(* IEC 61131-3 sources: TetherPLC/compat/tc3 (part 2) *)

(* ---- tc3_analytics.st ---- *)
// tc3_analytics.st — Tc3_Analytics surface (TF3510/TF3500/TF3520):
// measurement analytics.  TwinCAT's full library is ~670 APIs
// behind a licensed analytics engine; the local measurement-side
// primitives (event counting, windowed statistics, sample
// logging) are pure-ST here and fully functional, while the
// engine-backed surfaces (storage provider, MQTT/HTTP egress
// transport) report an honest engine-absent error.
//
// Differences from the TwinCAT library
// (docs/plc/compat/README.md):
//   - TwinCAT's class/method/object model is flattened into
//     FB_* blocks with Execute-style inputs, matching the other
//     TetherPLC compat surfaces.
//   - The ring logger exposes the newest N samples via indexed
//     outputs Slot0..Slot7 plus Count; a real circular-buffer
//     API needs dynamic memory we do not model.
//   - Storage/provider and transport FBs accept the command,
//     run a bounded handshake, then fail ErrorId=1
//     (engine-unavailable): no database or MQTT egress is faked.

// ---- FB_AnalyticsCounter: edge counter + rate per window ----
FUNCTION_BLOCK FB_AnalyticsCounter
VAR_INPUT
    Enable : BOOL;
    Event : BOOL;               // count rising edges
    WindowTime : LREAL;         // seconds per rate window
    CycleTime : LREAL;          // task cycle seconds
    Reset : BOOL;
END_VAR
VAR_OUTPUT
    Total : UDINT;
    WindowCount : UDINT;
    Rate : LREAL;               // events per second (last window)
    WindowDone : BOOL;
END_VAR
VAR
    prev : BOOL;
    acc : LREAL;
END_VAR
    WindowDone := FALSE;
    IF Reset THEN
        Total := 0;
        WindowCount := 0;
        Rate := 0.0;
        acc := 0.0;
        prev := FALSE;
    END_IF;
    IF NOT Enable THEN
        prev := Event;
        RETURN;
    END_IF;
    IF Event AND NOT prev THEN
        Total := Total + 1;
        WindowCount := WindowCount + 1;
    END_IF;
    prev := Event;
    acc := acc + CycleTime;
    IF WindowTime > 0.0 AND acc >= WindowTime THEN
        Rate := UDINT_TO_LREAL(WindowCount) / acc;
        WindowCount := 0;
        acc := 0.0;
        WindowDone := TRUE;
    END_IF;
END_FUNCTION_BLOCK

// ---- FB_AnalyticsStats: running + windowed min/max/mean ----
FUNCTION_BLOCK FB_AnalyticsStats
VAR_INPUT
    Execute : BOOL;             // sample the input when TRUE
    Sample : LREAL;
    Clear : BOOL;
END_VAR
VAR_OUTPUT
    Count : UDINT;
    Min : LREAL;
    Max : LREAL;
    Mean : LREAL;
    Valid : BOOL;
END_VAR
VAR
    sum : LREAL;
END_VAR
    Valid := FALSE;
    IF Clear THEN
        Count := 0;
        Min := 0.0;
        Max := 0.0;
        Mean := 0.0;
        sum := 0.0;
    END_IF;
    IF NOT Execute THEN RETURN; END_IF;
    IF Count = 0 THEN
        Min := Sample;
        Max := Sample;
    ELSE
        IF Sample < Min THEN Min := Sample; END_IF;
        IF Sample > Max THEN Max := Sample; END_IF;
    END_IF;
    Count := Count + 1;
    sum := sum + Sample;
    Mean := sum / UDINT_TO_LREAL(Count);
    Valid := TRUE;
END_FUNCTION_BLOCK

// ---- FB_AnalyticsLogger: 8-deep ring of timestamped samples ----
FUNCTION_BLOCK FB_AnalyticsLogger
VAR_INPUT
    Record : BOOL;              // rising edge stores a sample
    Value : LREAL;
    Timestamp : LREAL;          // caller-supplied time tag
    Clear : BOOL;
END_VAR
VAR_OUTPUT
    Count : UDINT;              // total records stored
    Slot0 : LREAL; Slot1 : LREAL; Slot2 : LREAL; Slot3 : LREAL;
    Slot4 : LREAL; Slot5 : LREAL; Slot6 : LREAL; Slot7 : LREAL;
    LastTs : LREAL;
    Overflow : BOOL;            // wrapped at least once
END_VAR
VAR
    head : UDINT;
    prev : BOOL;
END_VAR
    IF Clear THEN
        Count := 0;
        head := 0;
        LastTs := 0.0;
        Overflow := FALSE;
        Slot0 := 0.0; Slot1 := 0.0; Slot2 := 0.0; Slot3 := 0.0;
        Slot4 := 0.0; Slot5 := 0.0; Slot6 := 0.0; Slot7 := 0.0;
    END_IF;
    IF Record AND NOT prev THEN
        IF head = 0 THEN Slot0 := Value; END_IF;
        IF head = 1 THEN Slot1 := Value; END_IF;
        IF head = 2 THEN Slot2 := Value; END_IF;
        IF head = 3 THEN Slot3 := Value; END_IF;
        IF head = 4 THEN Slot4 := Value; END_IF;
        IF head = 5 THEN Slot5 := Value; END_IF;
        IF head = 6 THEN Slot6 := Value; END_IF;
        IF head = 7 THEN Slot7 := Value; END_IF;
        head := head + 1;
        IF head >= 8 THEN
            head := 0;
            Overflow := TRUE;
        END_IF;
        Count := Count + 1;
        LastTs := Timestamp;
    END_IF;
    prev := Record;
END_FUNCTION_BLOCK

// ---- FB_AnalyticsStore: engine-backed storage provider ----
// Honest engine-absent block: accepts a flush/store command,
// holds Busy for a bounded handshake, then fails with
// ErrorId=1 — no database write is ever claimed.
FUNCTION_BLOCK FB_AnalyticsStore
VAR_INPUT
    Execute : BOOL;
    Abort : BOOL;
    ProviderPath : STRING;      // e.g. database/Influx endpoint
    RecordCount : UDINT;
END_VAR
VAR_OUTPUT
    Busy : BOOL;
    Error : BOOL;
    ErrorId : UDINT;            // 0 none, 1 engine-unavailable,
                                // 2 bad-provider, 3 aborted
    Done : BOOL;
END_VAR
VAR
    phase : INT;
    tmo : UDINT;
END_VAR
    Done := FALSE;
    IF phase = 0 THEN
        Busy := FALSE;
        IF Execute THEN
            Busy := TRUE;
            Error := FALSE;
            ErrorId := 0;
            tmo := 0;
            IF ProviderPath = '' THEN
                Error := TRUE;
                ErrorId := 2;
                phase := 2;
            ELSE
                phase := 1;
            END_IF;
        END_IF;
    ELSIF phase = 1 THEN
        tmo := tmo + 1;
        IF tmo >= 4 THEN
            Busy := FALSE;
            Error := TRUE;
            ErrorId := 1;       // engine-unavailable
            phase := 2;
        END_IF;
    ELSE
        Busy := FALSE;
        IF NOT Execute THEN phase := 0; END_IF;
    END_IF;
    IF Abort AND phase = 1 THEN
        Busy := FALSE;
        Error := TRUE;
        ErrorId := 3;
        phase := 2;
    END_IF;
    Done := (phase = 2);
END_FUNCTION_BLOCK

(* ---- tc3_ba_common.st ---- *)
// tc3_ba_common.st — Tc3_BA_Common + Tc3_BA2_Common surface
// (TwinCAT_3_PLC_Lib_Tc3_BA*_Common_EN): pure-ST building-
// automation commons — time-of-day helpers, edge/COV triggers,
// ramp limiters, 2-point switches, PID, sequence controller,
// and a bounded dynamic array.  KL32xx terminal config is not
// modeled (blocks take scaled process values).
//
// Differences: the BA_* enum-validity helpers map to plain
// range checks (enums are INT here); the DynamicArray is a
// bounded fixed-capacity variant (no heap growth).

// ---- F_BA_RemMsTp: ms remaining to a target time ----
FUNCTION F_BA_RemMsTp : UDINT
VAR_INPUT
    tNow : UDINT;               // ms
    tTarget : UDINT;
END_VAR
    IF tTarget >= tNow THEN
        F_BA_RemMsTp := tTarget - tNow;
    ELSE
        F_BA_RemMsTp := 0;
    END_IF;
END_FUNCTION

// ---- F_BA_RemSecsTp: s remaining to a target ----
FUNCTION F_BA_RemSecsTp : UDINT
VAR_INPUT
    tNow : UDINT;
    tTarget : UDINT;
END_VAR
    IF tTarget >= tNow THEN
        F_BA_RemSecsTp := tTarget - tNow;
    ELSE
        F_BA_RemSecsTp := 0;
    END_IF;
END_FUNCTION

// ---- F_BA_IsWeekdayValid: 1..7 range check ----
FUNCTION F_BA_IsWeekdayValid : BOOL
VAR_INPUT
    day : INT;
END_VAR
    F_BA_IsWeekdayValid := day >= 1 AND day <= 7;
END_FUNCTION

// ---- F_BA_IsUnitValid: unit-id range check ----
FUNCTION F_BA_IsUnitValid : BOOL
VAR_INPUT
    unit : INT;
END_VAR
    F_BA_IsUnitValid := unit >= 0 AND unit <= 255;
END_FUNCTION

// ---- FB_BA_RFTrig: rising/falling edge detector ----
FUNCTION_BLOCK FB_BA_RFTrig
VAR_INPUT
    bIn : BOOL;
END_VAR
VAR_OUTPUT
    bRise : BOOL;
    bFall : BOOL;
END_VAR
VAR
    prev : BOOL;
END_VAR
    bRise := bIn AND NOT prev;
    bFall := NOT bIn AND prev;
    prev := bIn;
END_FUNCTION_BLOCK

// ---- FB_BA_ATrigCOV: change-of-value trigger ----
// Fires when the input changes by more than fDelta since the
// last reported value.
FUNCTION_BLOCK FB_BA_ATrigCOV
VAR_INPUT
    bEnable : BOOL;
    fIn : LREAL;
    fDelta : LREAL;
END_VAR
VAR_OUTPUT
    bTrig : BOOL;
    fOut : LREAL;
END_VAR
VAR
    fLast : LREAL;
    init : BOOL;
END_VAR
    bTrig := FALSE;
    IF NOT bEnable THEN init := FALSE; RETURN; END_IF;
    IF NOT init THEN
        fLast := fIn;
        init := TRUE;
        bTrig := TRUE;
        fOut := fIn;
        RETURN;
    END_IF;
    IF fIn - fLast >= fDelta OR fLast - fIn >= fDelta THEN
        fLast := fIn;
        fOut := fIn;
        bTrig := TRUE;
    END_IF;
END_FUNCTION_BLOCK

// ---- FB_BA_RampLmt: ramp with output clamp ----
FUNCTION_BLOCK FB_BA_RampLmt
VAR_INPUT
    bEnable : BOOL;
    fIn : LREAL;
    fSlewUp : LREAL;            // unit/s
    fSlewDown : LREAL;
    fMin : LREAL;
    fMax : LREAL;
    CycleTime : LREAL;
END_VAR
VAR_OUTPUT
    fOut : LREAL;
    bAtTarget : BOOL;
END_VAR
    IF NOT bEnable THEN bAtTarget := FALSE; RETURN; END_IF;
    IF fOut < fIn THEN
        fOut := fOut + fSlewUp * CycleTime;
        IF fOut > fIn THEN fOut := fIn; END_IF;
    ELSIF fOut > fIn THEN
        fOut := fOut - fSlewDown * CycleTime;
        IF fOut < fIn THEN fOut := fIn; END_IF;
    END_IF;
    IF fOut > fMax THEN fOut := fMax; END_IF;
    IF fOut < fMin THEN fOut := fMin; END_IF;
    bAtTarget := fOut = fIn;
END_FUNCTION_BLOCK

// ---- FB_BA_Swi2P: two-point switch ----
FUNCTION_BLOCK FB_BA_Swi2P
VAR_INPUT
    bEnable : BOOL;
    fIn : LREAL;
    fOn : LREAL;
    fOff : LREAL;
END_VAR
VAR_OUTPUT
    bOut : BOOL;
END_VAR
VAR
    q : BOOL;
END_VAR
    IF NOT bEnable THEN q := FALSE; bOut := FALSE; RETURN; END_IF;
    IF fIn >= fOn THEN q := TRUE; END_IF;
    IF fIn <= fOff THEN q := FALSE; END_IF;
    bOut := q;
END_FUNCTION_BLOCK

// ---- FB_BA_SwiHys2P: two-point switch with hysteresis ----
FUNCTION_BLOCK FB_BA_SwiHys2P
VAR_INPUT
    bEnable : BOOL;
    fIn : LREAL;
    fSp : LREAL;
    fHys : LREAL;
    bInvert : BOOL;
END_VAR
VAR_OUTPUT
    bOut : BOOL;
END_VAR
VAR
    q : BOOL;
END_VAR
    IF NOT bEnable THEN q := FALSE; bOut := FALSE; RETURN; END_IF;
    IF bInvert THEN
        IF fIn >= fSp + fHys THEN q := TRUE; END_IF;
        IF fIn <= fSp THEN q := FALSE; END_IF;
    ELSE
        IF fIn <= fSp - fHys THEN q := TRUE; END_IF;
        IF fIn >= fSp THEN q := FALSE; END_IF;
    END_IF;
    bOut := q;
END_FUNCTION_BLOCK

// ---- FB_BA_PIDCtrl: PI controller with anti-windup ----
FUNCTION_BLOCK FB_BA_PIDCtrl
VAR_INPUT
    bEnable : BOOL;
    fActual : LREAL;
    fSetpoint : LREAL;
    fKp : LREAL;
    fTi : LREAL;                // s; 0 = P only
    fOutMin : LREAL;
    fOutMax : LREAL;
    CycleTime : LREAL;
END_VAR
VAR_OUTPUT
    fOut : LREAL;
    fError : LREAL;
END_VAR
VAR
    iTerm : LREAL;
END_VAR
    IF NOT bEnable THEN
        fOut := fOutMin; iTerm := 0.0; fError := 0.0;
        RETURN;
    END_IF;
    fError := fSetpoint - fActual;
    iTerm := iTerm + fError * CycleTime;
    fOut := fKp * fError;
    IF fTi > 0.0 THEN
        fOut := fKp * (fError + iTerm / fTi);
    END_IF;
    IF fOut > fOutMax THEN
        fOut := fOutMax;
        iTerm := iTerm - fError * CycleTime;
    END_IF;
    IF fOut < fOutMin THEN
        fOut := fOutMin;
        iTerm := iTerm - fError * CycleTime;
    END_IF;
END_FUNCTION_BLOCK

// ---- FB_BA_SeqCtrl: sequence controller ----
// Distributes a 0..100 demand across up to 4 sequential
// stages (each stage gets a slice of the demand range).
FUNCTION_BLOCK FB_BA_SeqCtrl
VAR_INPUT
    bEnable : BOOL;
    fDemand : LREAL;            // 0..100 %
    nStages : INT;              // 1..4
END_VAR
VAR_OUTPUT
    fStage1 : LREAL;            // each 0..100
    fStage2 : LREAL;
    fStage3 : LREAL;
    fStage4 : LREAL;
END_VAR
VAR
    seg : LREAL;
    rem : LREAL;
    nR : LREAL;
END_VAR
    IF NOT bEnable OR nStages <= 0 THEN
        fStage1 := 0.0; fStage2 := 0.0;
        fStage3 := 0.0; fStage4 := 0.0;
        RETURN;
    END_IF;
    nR := DINT_TO_LREAL(INT_TO_DINT(nStages));
    seg := 100.0 / nR;
    rem := fDemand;
    fStage1 := rem; IF fStage1 > seg THEN fStage1 := seg; END_IF;
    IF fStage1 < 0.0 THEN fStage1 := 0.0; END_IF;
    rem := rem - seg;
    fStage2 := rem; IF fStage2 > seg THEN fStage2 := seg; END_IF;
    IF fStage2 < 0.0 THEN fStage2 := 0.0; END_IF;
    rem := rem - seg;
    fStage3 := rem; IF fStage3 > seg THEN fStage3 := seg; END_IF;
    IF fStage3 < 0.0 THEN fStage3 := 0.0; END_IF;
    rem := rem - seg;
    fStage4 := rem; IF fStage4 > seg THEN fStage4 := seg; END_IF;
    IF fStage4 < 0.0 THEN fStage4 := 0.0; END_IF;
    // normalize each stage to 0..100 of its own slice
    fStage1 := fStage1 * 100.0 / seg;
    fStage2 := fStage2 * 100.0 / seg;
    fStage3 := fStage3 * 100.0 / seg;
    fStage4 := fStage4 * 100.0 / seg;
END_FUNCTION_BLOCK

// ---- FB_BA_DynamicArray: bounded key->value store ----
// Fixed capacity 16; key 0 is empty.
FUNCTION_BLOCK FB_BA_DynamicArray
VAR_INPUT
    bEnable : BOOL;
    Op : INT;                   // 1=set, 2=get, 3=remove, 4=find
    Key : UDINT;
    Value : LREAL;
END_VAR
VAR_OUTPUT
    Done : BOOL;
    Found : BOOL;
    OutValue : LREAL;
    Count : INT;
    Free : INT;
END_VAR
VAR
    keys : ARRAY[0..15] OF UDINT;
    vals : ARRAY[0..15] OF LREAL;
    cnt : INT;
    i : INT;
    slot : INT;
END_VAR
    Done := FALSE;
    Found := FALSE;
    OutValue := 0.0;
    IF NOT bEnable THEN RETURN; END_IF;
    slot := -1;
    FOR i := 0 TO 15 DO
        IF keys[i] = Key THEN slot := i; END_IF;
    END_FOR;
    IF Op = 1 THEN
        IF slot >= 0 THEN
            vals[slot] := Value;
            Found := TRUE;
            Done := TRUE;
        ELSE
            FOR i := 0 TO 15 DO
                IF slot < 0 AND keys[i] = 0 THEN slot := i; END_IF;
            END_FOR;
            IF slot >= 0 THEN
                keys[slot] := Key;
                vals[slot] := Value;
                cnt := cnt + 1;
                Done := TRUE;
            END_IF;
        END_IF;
    ELSIF Op = 2 OR Op = 4 THEN
        IF slot >= 0 THEN
            Found := TRUE;
            Done := TRUE;
            OutValue := vals[slot];
        END_IF;
    ELSIF Op = 3 THEN
        IF slot >= 0 THEN
            keys[slot] := 0;
            vals[slot] := 0.0;
            cnt := cnt - 1;
            Found := TRUE;
            Done := TRUE;
        END_IF;
    END_IF;
    Count := cnt;
    Free := 16 - cnt;
END_FUNCTION_BLOCK

(* ---- tc3_bacnet.st ---- *)
// Tc3_sACN -> Tc3_BACnetRev14 BACnet/IP client wrappers.
// Beckhoff's BACnet integration is device-configuration-driven
// (FBs are generated per configured device in TwinCAT), so there
// is no static TwinCAT FB API to mirror; these wrappers expose
// the tplc-bacnet service (ASHRAE 135 over UDP 47808) as
// poll-driven function blocks in the same shape as the other
// compat libraries.
// Differences from a TwinCAT BACnet device binding, documented in
// docs/plc/compat/README.md:
//   - Who-Is/ReadProperty/WriteProperty only; no COV subscriptions,
//     no device-object discovery beyond I-Am fields, no segmentation.
//   - Values cross as raw BACnet application-tag payload bytes:
//     nValueType selects the tag (1=boolean, 2=unsigned, 3=integer,
//     4=real, 5=double, 6=octetString, 7=characterString,
//     9=enumerated, 12=objectIdentifier) and pValue holds the tag
//     payload in wire byte order.
//   - nErrId carries tplc-bacnet service/transport codes.
// Sources: docs/plc/plan/21-twincat-libraries.md §7 (TF8020).

FUNCTION_BLOCK FB_BACnet_WhoIs
VAR_INPUT
    sHost : STRING[15];        // "" or "255.255.255.255" = broadcast
    nPort : UDINT := 47808;
    bHasRange : BOOL;
    nRangeLo : UDINT;
    nRangeHi : UDINT;
    bExecute : BOOL;
    tTimeout : TIME := T#1S;
END_VAR
VAR_OUTPUT
    bBusy : BOOL;
    bDone : BOOL;
    bError : BOOL;
    nErrId : UDINT;
    nStatus : DINT;
    nDevCount : UDINT;
    nDevId : ARRAY[0..7] OF UDINT;   // (objType<<22)|instance
    nDevIp : ARRAY[0..31] OF BYTE;   // 4 bytes per device
    nDevVendor : UDINT;
    nDevMaxApdu : UDINT;
    nDevSeg : UDINT;
END_VAR
VAR
    bac : FB_Bacnet;
    i : UDINT;
END_VAR
    bac.FUNC := 1;
    bac.HOST := sHost;
    bac.PORT := nPort;
    bac.HAS_RANGE := bHasRange;
    bac.RANGE_LO := nRangeLo;
    bac.RANGE_HI := nRangeHi;
    bac.TIMEOUT := tTimeout;
    bac.EXEC := bExecute;
    bac();
    bBusy := bac.BUSY;
    bDone := bac.DONE;
    nStatus := bac.STATUS;
    nErrId := bac.ERRID;
    nDevCount := bac.DEV_COUNT;
    nDevVendor := bac.DEV_VENDOR;
    nDevMaxApdu := bac.DEV_MAX_APDU;
    nDevSeg := bac.DEV_SEG;
    IF bac.DONE THEN
        i := 0;
        WHILE i < bac.DEV_COUNT AND i < 8 DO
            nDevId[i] := bac.DEV_ID[i];
            nDevIp[i*4] := bac.DEV_IP[i*4];
            nDevIp[i*4+1] := bac.DEV_IP[i*4+1];
            nDevIp[i*4+2] := bac.DEV_IP[i*4+2];
            nDevIp[i*4+3] := bac.DEV_IP[i*4+3];
            i := i + 1;
        END_WHILE;
    END_IF;
    bError := (bac.ERRID <> 0) OR (bac.STATUS >= 2);
END_FUNCTION_BLOCK

FUNCTION_BLOCK FB_BACnet_ReadProperty
VAR_INPUT
    sHost : STRING[15];
    nPort : UDINT := 47808;
    nObjType : UDINT;          // e.g. 8=device, 0=analogInput
    nObjInst : UDINT;
    nPropId : UDINT;           // e.g. 85=present-value, 77=object-name
    bHasIdx : BOOL;
    nPropIdx : UDINT;          // array index when bHasIdx
    bExecute : BOOL;
    tTimeout : TIME := T#1S;
END_VAR
VAR_OUTPUT
    bBusy : BOOL;
    bDone : BOOL;
    bError : BOOL;
    nErrId : UDINT;
    nStatus : DINT;
    nService : UDINT;
    nApdu : UDINT;
    nRObjType : UDINT;
    nRObjInst : UDINT;
    nRPropId : UDINT;
    nValueType : UDINT;        // app tag of returned value
    nValueLen : UDINT;
    pValue : ARRAY[0..255] OF BYTE;
END_VAR
VAR
    bac : FB_Bacnet;
    i : UDINT;
END_VAR
    bac.FUNC := 2;
    bac.HOST := sHost;
    bac.PORT := nPort;
    bac.OBJ_TYPE := nObjType;
    bac.OBJ_INST := nObjInst;
    bac.PROP_ID := nPropId;
    bac.HAS_IDX := bHasIdx;
    bac.PROP_IDX := nPropIdx;
    bac.TIMEOUT := tTimeout;
    bac.EXEC := bExecute;
    bac();
    bBusy := bac.BUSY;
    bDone := bac.DONE;
    nStatus := bac.STATUS;
    nErrId := bac.ERRID;
    nService := bac.R_SERVICE;
    nApdu := bac.R_APDU;
    nRObjType := bac.R_OBJ_TYPE;
    nRObjInst := bac.R_OBJ_INST;
    nRPropId := bac.R_PROP_ID;
    nValueType := bac.R_VTYPE;
    nValueLen := bac.R_VLEN;
    IF bac.DONE THEN
        i := 0;
        WHILE i < bac.R_VLEN AND i < 256 DO
            pValue[i] := bac.R_VAL[i];
            i := i + 1;
        END_WHILE;
    END_IF;
    bError := (bac.ERRID <> 0) OR (bac.STATUS >= 2);
END_FUNCTION_BLOCK

FUNCTION_BLOCK FB_BACnet_WriteProperty
VAR_INPUT
    sHost : STRING[15];
    nPort : UDINT := 47808;
    nObjType : UDINT;
    nObjInst : UDINT;
    nPropId : UDINT;
    bHasIdx : BOOL;
    nPropIdx : UDINT;
    nValueType : UDINT;        // app tag for the value
    nValueLen : UDINT;
    pValue : ARRAY[0..255] OF BYTE;
    bHasPrio : BOOL;
    nPriority : UDINT;         // 1..16 when bHasPrio
    bExecute : BOOL;
    tTimeout : TIME := T#1S;
END_VAR
VAR_OUTPUT
    bBusy : BOOL;
    bDone : BOOL;
    bError : BOOL;
    nErrId : UDINT;
    nStatus : DINT;
    nService : UDINT;
END_VAR
VAR
    bac : FB_Bacnet;
    i : UDINT;
END_VAR
    bac.FUNC := 3;
    bac.HOST := sHost;
    bac.PORT := nPort;
    bac.OBJ_TYPE := nObjType;
    bac.OBJ_INST := nObjInst;
    bac.PROP_ID := nPropId;
    bac.HAS_IDX := bHasIdx;
    bac.PROP_IDX := nPropIdx;
    bac.VAL_TYPE := nValueType;
    bac.VLEN := nValueLen;
    i := 0;
    WHILE i < nValueLen AND i < 256 DO
        bac.VAL[i] := pValue[i];
        i := i + 1;
    END_WHILE;
    bac.HAS_PRIO := bHasPrio;
    bac.PRIORITY := nPriority;
    bac.TIMEOUT := tTimeout;
    bac.EXEC := bExecute;
    bac();
    bBusy := bac.BUSY;
    bDone := bac.DONE;
    nStatus := bac.STATUS;
    nErrId := bac.ERRID;
    nService := bac.R_SERVICE;
    bError := (bac.ERRID <> 0) OR (bac.STATUS >= 2);
END_FUNCTION_BLOCK

(* ---- tc3_database.st ---- *)
// Tc2_Database / Tc3_Database -> SQL surface over the tplc-db
// service (embedded SQLite, no TwinCAT Database Server, no
// ODBC driver manager).  Documented differences:
//   - Statements are plain SQL text (SQLite dialect).
//   - Query results cross as tab-separated rows in a bounded
//     255-byte buffer; ROWS/COLS report the produced shape.
//   - METHOD calls are edge-triggered command inputs (nCmd).
//   - The TF6420 configuration/AutoLog/event families
//     (FB_ConfigTcDBSrvEvt, FB_PLCDBAutoLogEvt) are not
//     modelled; the PLC DB access blocks are.
//   - nErrId carries tplc-db service codes; GetError returns the
//     engine's last error text.

// ---- FB_PLCDBOpen: open/create a database ----
FUNCTION_BLOCK FB_PLCDBOpen
VAR_INPUT
    nCmd : UDINT;               // 1 open, 4 close
    sPath : STRING[127];
END_VAR
VAR_OUTPUT
    hDb : UDINT;
    bDone : BOOL;
    bBusy : BOOL;
    bError : BOOL;
    nErrId : UDINT;
END_VAR
VAR
    db : FB_Db;
    prev : UDINT;
END_VAR
    bDone := FALSE; bError := FALSE; nErrId := 0; bBusy := FALSE;
    IF nCmd <> 0 AND prev = 0 THEN
        bBusy := TRUE;
        db.OP := nCmd;
        db.HANDLE := hDb;
        db.PATH := sPath;
        db();
        bBusy := FALSE;
        IF db.STATUS = 0 THEN
            bDone := TRUE;
            IF nCmd = 1 THEN hDb := db.HANDLE; ELSE hDb := 0; END_IF;
        ELSE
            bError := TRUE; nErrId := db.ERRID;
        END_IF;
    END_IF;
    prev := nCmd;
END_FUNCTION_BLOCK

// ---- FB_PLCDBCreateEvt: CREATE/DDL and other exec statements ----
FUNCTION_BLOCK FB_PLCDBCreateEvt
VAR_INPUT
    nCmd : UDINT;               // 2 exec
    hDb : UDINT;
    sSql : STRING[255];
END_VAR
VAR_OUTPUT
    nChanges : UDINT;
    bDone : BOOL;
    bBusy : BOOL;
    bError : BOOL;
    nErrId : UDINT;
END_VAR
VAR
    db : FB_Db;
    prev : UDINT;
END_VAR
    bDone := FALSE; bError := FALSE; nErrId := 0; bBusy := FALSE;
    IF nCmd <> 0 AND prev = 0 THEN
        bBusy := TRUE;
        db.OP := 2; db.HANDLE := hDb; db.SQL := sSql;
        db();
        bBusy := FALSE;
        IF db.STATUS = 0 THEN
            bDone := TRUE; nChanges := db.CHANGES;
        ELSE
            bError := TRUE; nErrId := db.ERRID;
        END_IF;
    END_IF;
    prev := nCmd;
END_FUNCTION_BLOCK

// ---- FB_PLCDBWriteEvt: INSERT/UPDATE/DELETE ----
FUNCTION_BLOCK FB_PLCDBWriteEvt
VAR_INPUT
    nCmd : UDINT;               // 2 exec
    hDb : UDINT;
    sSql : STRING[255];
END_VAR
VAR_OUTPUT
    nChanges : UDINT;
    bDone : BOOL;
    bBusy : BOOL;
    bError : BOOL;
    nErrId : UDINT;
END_VAR
VAR
    db : FB_Db;
    prev : UDINT;
END_VAR
    bDone := FALSE; bError := FALSE; nErrId := 0; bBusy := FALSE;
    IF nCmd <> 0 AND prev = 0 THEN
        bBusy := TRUE;
        db.OP := 2; db.HANDLE := hDb; db.SQL := sSql;
        db();
        bBusy := FALSE;
        IF db.STATUS = 0 THEN
            bDone := TRUE; nChanges := db.CHANGES;
        ELSE
            bError := TRUE; nErrId := db.ERRID;
        END_IF;
    END_IF;
    prev := nCmd;
END_FUNCTION_BLOCK

// ---- FB_PLCDBReadEvt: SELECT -> rows/cols + text buffer ----
FUNCTION_BLOCK FB_PLCDBReadEvt
VAR_INPUT
    nCmd : UDINT;               // 3 query
    hDb : UDINT;
    sSql : STRING[255];
END_VAR
VAR_OUTPUT
    nRows : UDINT;
    nCols : UDINT;
    sResult : STRING[255];      // tab-separated, '\n' per row
    bDone : BOOL;
    bBusy : BOOL;
    bError : BOOL;
    nErrId : UDINT;
END_VAR
VAR
    db : FB_Db;
    prev : UDINT;
END_VAR
    bDone := FALSE; bError := FALSE; nErrId := 0; bBusy := FALSE;
    IF nCmd <> 0 AND prev = 0 THEN
        bBusy := TRUE;
        db.OP := 3; db.HANDLE := hDb; db.SQL := sSql;
        db();
        bBusy := FALSE;
        IF db.STATUS = 0 THEN
            bDone := TRUE;
            nRows := db.ROWS; nCols := db.COLS;
            sResult := db.BUF;
        ELSE
            bError := TRUE; nErrId := db.ERRID;
        END_IF;
    END_IF;
    prev := nCmd;
END_FUNCTION_BLOCK

// ---- FB_PLCDBGetError: engine error text ----
FUNCTION_BLOCK FB_PLCDBGetError
VAR_INPUT
    nCmd : UDINT;               // 5 error
    hDb : UDINT;
END_VAR
VAR_OUTPUT
    sError : STRING[127];
    bDone : BOOL;
    bError : BOOL;
    nErrId : UDINT;
END_VAR
VAR
    db : FB_Db;
    prev : UDINT;
END_VAR
    bDone := FALSE; bError := FALSE; nErrId := 0;
    IF nCmd <> 0 AND prev = 0 THEN
        db.OP := 5; db.HANDLE := hDb;
        db();
        IF db.STATUS = 0 THEN
            bDone := TRUE; sError := db.ERR;
        ELSE
            bError := TRUE; nErrId := db.ERRID;
        END_IF;
    END_IF;
    prev := nCmd;
END_FUNCTION_BLOCK

(* ---- tc3_dynmem.st ---- *)
// Tc3_DynamicMemory -> FB_DynMem_Buffer / FB_DynMem_Manager.
// Beckhoff's originals hand out PVOIDs into a shared heap; we
// model the same behaviour over the tplc-dynmem bounded arena —
// blocks are integer handles (never raw pointers), accessed via
// FB_DynMem_Access byte I/O.  Documented differences:
//   - No POINTER semantics: a "buffer" is a handle; data crosses
//     one byte at a time through FB_DynMem_Access.
//   - METHOD calls are expressed as edge-triggered command
//     inputs (this compiler has no METHOD support): nCmd
//     1=Allocate 2=Reallocate 3=Deallocate.
//   - Arena is fixed (64 blocks, 64 KiB max block, 1 MiB total)
//     — deterministic worst case, no host-heap interaction.
//   - nErrId carries tplc-dynmem service codes.

// ---- FB_DynMem_Buffer: owned buffer handle ----
FUNCTION_BLOCK FB_DynMem_Buffer
VAR_INPUT
    nCmd : UDINT;               // 0 none, 1 alloc, 2 realloc, 3 dealloc
    nNewSize : UDINT;
    bPreserve : BOOL;
    bReset : BOOL;
END_VAR
VAR_OUTPUT
    hBuffer : UDINT;            // 0 = not allocated
    nSize : UDINT;
    bDone : BOOL;
    bError : BOOL;
    nErrId : UDINT;
END_VAR
VAR
    dm : FB_DynMem;
    prev : UDINT;
END_VAR
    bDone := FALSE; bError := FALSE; nErrId := 0;
    IF nCmd <> 0 AND prev = 0 THEN
        IF nCmd = 1 THEN
            dm.OP := 1; dm.SIZE := nNewSize;
            dm.RESET := BOOL_TO_UDINT(bReset);
        ELSIF nCmd = 2 THEN
            IF hBuffer = 0 THEN
                bError := TRUE; nErrId := 2;
            ELSE
                dm.OP := 3; dm.ID := hBuffer; dm.SIZE := nNewSize;
                dm.PRESERVE := BOOL_TO_UDINT(bPreserve);
                dm.RESET := BOOL_TO_UDINT(bReset);
            END_IF;
        ELSIF nCmd = 3 THEN
            dm.OP := 2; dm.ID := hBuffer;
        END_IF;
        IF NOT bError THEN
            dm();
            IF dm.STATUS = 0 THEN
                bDone := TRUE;
                IF nCmd = 1 THEN
                    hBuffer := dm.ID; nSize := nNewSize;
                ELSIF nCmd = 2 THEN
                    nSize := nNewSize;
                ELSE
                    hBuffer := 0; nSize := 0;
                END_IF;
            ELSE
                bError := TRUE; nErrId := dm.ERRID;
            END_IF;
        END_IF;
    END_IF;
    prev := nCmd;
END_FUNCTION_BLOCK

// ---- FB_DynMem_Access: byte I/O into a block handle ----
FUNCTION_BLOCK FB_DynMem_Access
VAR_INPUT
    nCmd : UDINT;               // 0 none, 4 read, 5 write
    nHandle : UDINT;
    nOffset : UDINT;
    nByte : BYTE;
END_VAR
VAR_OUTPUT
    nOut : BYTE;
    bDone : BOOL;
    bError : BOOL;
    nErrId : UDINT;
END_VAR
VAR
    dm : FB_DynMem;
    prev : UDINT;
END_VAR
    bDone := FALSE; bError := FALSE; nErrId := 0;
    IF nCmd <> 0 AND prev = 0 THEN
        IF nCmd = 4 OR nCmd = 5 THEN
            dm.OP := nCmd; dm.ID := nHandle; dm.OFFSET := nOffset;
            dm.BYTE := BYTE_TO_UDINT(nByte);
            dm();
            IF dm.STATUS = 0 THEN
                bDone := TRUE;
                IF nCmd = 4 THEN nOut := UDINT_TO_BYTE(dm.BYTE); END_IF;
            ELSE
                bError := TRUE; nErrId := dm.ERRID;
            END_IF;
        END_IF;
    END_IF;
    prev := nCmd;
END_FUNCTION_BLOCK

// ---- FB_DynMem_Manager: alloc/free + consumption counters ----
FUNCTION_BLOCK FB_DynMem_Manager
VAR_INPUT
    nCmd : UDINT;               // 0 none, 1 alloc, 3 dealloc
    nReqSize : UDINT;
    bReset : BOOL;
    nId : UDINT;                // dealloc target
END_VAR
VAR_OUTPUT
    hNew : UDINT;               // handle returned by alloc
    bDone : BOOL;
    bError : BOOL;
    nErrId : UDINT;
    nLiveBlocks : UDINT;
    nLiveBytes : UDINT;
    nTotalAllocs : UDINT;
    nTotalFrees : UDINT;
    nArenaBytes : UDINT;
    nArenaUsed : UDINT;
END_VAR
VAR
    dm : FB_DynMem;
    prev : UDINT;
END_VAR
    bDone := FALSE; bError := FALSE; nErrId := 0;
    IF nCmd <> 0 AND prev = 0 THEN
        IF nCmd = 1 THEN
            dm.OP := 1; dm.SIZE := nReqSize;
            dm.RESET := BOOL_TO_UDINT(bReset);
            dm();
            IF dm.STATUS = 0 THEN
                bDone := TRUE; hNew := dm.ID;
            ELSE
                bError := TRUE; nErrId := dm.ERRID;
            END_IF;
        ELSIF nCmd = 3 THEN
            dm.OP := 2; dm.ID := nId;
            dm();
            IF dm.STATUS = 0 THEN
                bDone := TRUE;
            ELSE
                bError := TRUE; nErrId := dm.ERRID;
            END_IF;
        END_IF;
    END_IF;
    prev := nCmd;
    // refresh counters every invocation
    dm.OP := 6;
    dm();
    IF dm.STATUS = 0 THEN
        nLiveBlocks := dm.LIVEBLKS;
        nLiveBytes := dm.LIVEBYTES;
        nTotalAllocs := dm.TOTALALLOCS;
        nTotalFrees := dm.TOTALFREES;
        nArenaBytes := dm.ARENABYTES;
        nArenaUsed := dm.ARENAUSED;
    END_IF;
END_FUNCTION_BLOCK

(* ---- tc3_ecdiag.st ---- *)
// tc3_ecdiag.st — Tc3_EtherCATDiag compatibility surface.
//
// TwinCAT's EtherCAT diagnostics library reads the CoE 0x10F3
// "Diagnosis History" object from EtherCAT slaves.  TetherPLC bridges
// this onto the tplc-ecdiag host service, which reads the
// ec.coediag.* params exposed by a Tether IO endpoint
// (tether_io_motion_server in sim mode; a real master would bridge
// per-slave SDO reads of 0x10F3 under the same names).
//
// FB_EcDiagRead (builtin, layout FB_EcDiagRead):
//   OP      1 = read history, 2 = acknowledge (ACKVAL = newest acked)
//   SLAVE   slave port address
//   outputs COUNT NEWEST ACKED NEWMSGS INFOFLAGS STATUS ERRID plus
//           16-slot parallel entry arrays MSGTYPE ACKST TSMS CODE
//           CODETYPE TEXTID MODULE CHANNEL MSGTEXT
// STATUS is the service return code (0 ok, negative error), ERRID
// its positive magnitude.  When the service is inactive STATUS = -2.
//
// Mapping notes (documented deviations from the TwinCAT surface):
//   - ST_CoE_DiagHistory_Entry is a TwinCAT STRUCT; this dialect has
//     no user STRUCTs, so entries are exposed as parallel member
//     arrays aE* on FB_CoE_DiagHistory_Read (slot i = entry i).
//   - stTimeStamp TIMESTRUCT is flattened to aETimestampMs (ms since
//     the slave timestamp epoch reported by the device).
//   - sMsgText carries a generated "TID=/CODE=" string; real message
//     texts come from the slave ESI/XML which is not available.
//   - tReadInterval is approximated by nReadIntervalScans (scan
//     count, not wall time) since the scan period is not visible to
//     the FB.
//   - FB_CoE_DiagHistory_ReadAxis (AXIS_REF variant) is not provided:
//     it needs Tc2_MC2 axis objects; use the address variant.
//   - diag_code_type is approximated (emergency flag -> Emergency,
//     nonzero code -> DeviceRelated); module/profile typing needs
//     device profile data.
//
// SPDX-License-Identifier: Apache-2.0 OR MPL-2.0

// ---- FB_CoE_DiagHistory_Read -------------------------------------
// bEnable: rising edge reads once; while held, re-reads every
// nReadIntervalScans calls.  bAck (rising edge) acknowledges all
// messages up to NEWEST, then triggers a fresh read.

FUNCTION_BLOCK FB_CoE_DiagHistory_Read
VAR_INPUT
    sNetId : STRING[22];          // T_AmsNetId (accepted, unused)
    nSlaveAddr : UINT;            // slave port address
    bEnable : BOOL;
    bAck : BOOL;
    tTimeout : TIME := T#5S;      // accepted; IO is internally bounded
    tReadInterval : TIME := T#10S;// accepted; see nReadIntervalScans
    nReadIntervalScans : UDINT := 1000;
    // ST_CoE_DiagHistory_Options (flattened)
    nLangId : DINT := 1033;
    eBufferMode : USINT := 0;
    bEnableEmergSending : BOOL := TRUE;
    bFilterOutInfoMsgs : BOOL := FALSE;
    bFilterOutWarnMsgs : BOOL := FALSE;
    bFilterOutErrMsgs : BOOL := FALSE;
    bDisableAutoRecoverAfterConnectionErr : BOOL := FALSE;
    bExcludeTextIdFromMsgText : BOOL := FALSE;
END_VAR
VAR_OUTPUT
    bBusy : BOOL;
    bValid : BOOL;
    bError : BOOL;
    nErrorId : UDINT;
    // ST_CoE_DiagHistory_Info (flattened)
    bNewMsgsAvail : BOOL;
    bEmergSendingEnabled : BOOL;
    bInfoMsgsDisabled : BOOL;
    bWarnMsgsDisabled : BOOL;
    bErrMsgsDisabled : BOOL;
    bOldMsgsOverwritten : BOOL;
    bNewMsgsDiscarded : BOOL;
    // object header mirrors (sticky after each read)
    oNewest : UDINT;
    oAcked : UDINT;
    oNewMsgs : UDINT;
    oCount : UDINT;
END_VAR
VAR
    raw : FB_EcDiagRead;
    scanN : UDINT;
    prevEn : BOOL;
    prevAck : BOOL;
    haveResult : BOOL;
    lastOk : BOOL;
    i : UDINT;
    j : UDINT;
    keep : BOOL;
    // flattened entry arrays (public-readable member data)
    aEMsgType : ARRAY[0..15] OF UDINT;
    aEAckStatus : ARRAY[0..15] OF UDINT;
    aETimestampMs : ARRAY[0..15] OF UDINT;
    aEDiagCode : ARRAY[0..15] OF UDINT;
    aEDiagCodeType : ARRAY[0..15] OF UDINT;
    aETextId : ARRAY[0..15] OF UDINT;
    aEModuleNo : ARRAY[0..15] OF UDINT;
    aEChannelNo : ARRAY[0..15] OF UDINT;
    aEMsgText : ARRAY[0..15] OF STRING[63];
END_VAR
    bBusy := FALSE;
    bValid := haveResult AND lastOk;
    bError := haveResult AND NOT lastOk;
    nErrorId := 0;

    // acknowledge request: write newest as acked, then re-read below
    IF bAck AND NOT prevAck THEN
        raw.OP := 2;
        raw.SLAVE := nSlaveAddr;
        raw.ACKVAL := oNewest;
        raw();
        IF raw.STATUS < 0 THEN
            haveResult := TRUE;
            lastOk := FALSE;
            nErrorId := raw.ERRID;
        ELSE
            haveResult := TRUE;
            lastOk := TRUE;
        END_IF;
        scanN := 0;
    END_IF;

    // read trigger: rising edge, ack edge, or level-held interval
    IF (bEnable AND NOT prevEn) OR
       (bEnable AND scanN >= nReadIntervalScans) OR
       (bAck AND NOT prevAck) THEN
        raw.OP := 1;
        raw.SLAVE := nSlaveAddr;
        raw();
        bBusy := TRUE;   // service call is synchronous; pulses this scan
        haveResult := TRUE;
        lastOk := raw.STATUS >= 0;
        IF NOT lastOk THEN
            nErrorId := raw.ERRID;
        END_IF;
        scanN := 0;
    ELSIF bEnable THEN
        scanN := scanN + 1;
    END_IF;

    // mirror the object header (sticky across scans)
    oNewest := raw.NEWEST;
    oAcked := raw.ACKED;
    oNewMsgs := raw.NEWMSGS;
    oCount := raw.COUNT;

    // flatten raw entry arrays into the public aE* arrays, applying
    // the option filters (info/warn/error suppression)
    j := 0;
    FOR i := 0 TO 15 DO
        keep := i < raw.COUNT;
        IF keep AND bFilterOutInfoMsgs AND raw.MSGTYPE[i] = 1 THEN
            keep := FALSE;
        END_IF;
        IF keep AND bFilterOutWarnMsgs AND raw.MSGTYPE[i] = 2 THEN
            keep := FALSE;
        END_IF;
        IF keep AND bFilterOutErrMsgs AND raw.MSGTYPE[i] = 3 THEN
            keep := FALSE;
        END_IF;
        IF keep THEN
            aEMsgType[j] := raw.MSGTYPE[i];
            aEAckStatus[j] := raw.ACKST[i];
            aETimestampMs[j] := raw.TSMS[i];
            aEDiagCode[j] := raw.CODE[i];
            aEDiagCodeType[j] := raw.CODETYPE[i];
            aETextId[j] := raw.TEXTID[i];
            aEModuleNo[j] := raw.MODULE[i];
            aEChannelNo[j] := raw.CHANNEL[i];
            aEMsgText[j] := raw.MSGTEXT[i];
            j := j + 1;
        END_IF;
    END_FOR;

    // stInfo echo of the option inputs plus object state
    bNewMsgsAvail := oNewMsgs <> 0;
    bEmergSendingEnabled := bEnableEmergSending;
    bInfoMsgsDisabled := bFilterOutInfoMsgs;
    bWarnMsgsDisabled := bFilterOutWarnMsgs;
    bErrMsgsDisabled := bFilterOutErrMsgs;
    bOldMsgsOverwritten := FALSE;   // overwrite-mode tracking unsupported
    bNewMsgsDiscarded := FALSE;     // ack-mode discard tracking unsupported

    prevEn := bEnable;
    prevAck := bAck;
END_FUNCTION_BLOCK

(* ---- tc3_ecsync.st ---- *)
// tc3_ecsync.st — Tc3_EtherCATExtSync compatibility surface.
//
// TwinCAT's EtherCAT external-sync library exposes FBs that request
// and report the distributed-clock (DC) synchronization state of the
// EtherCAT master.  TetherPLC bridges those semantics onto the
// tplc-ecsync host service, which reads/writes the ec.dc.* params
// exposed by a Tether IO endpoint (tether_io_motion_server in sim
// mode, or a real master bridging DCManager/EtherCATDC stats under
// the same names).
//
// FB_EcSync (builtin, layout FB_EcSync):
//   OP      1 = poll status, 2 = set sync enable
//   ENABLE  sync enable value for OP 2 (0/1)
//   outputs CONNECTED SYNCEN PARAMSOK LASTERR STATUS ERRID DIFFNS
//           REFNS
// STATUS is the service return code (0 ok, negative error), ERRID
// its positive magnitude.  When the service is inactive (no
// TPLC_EC_IO/TPLC_MOTION_IO endpoint, or the endpoint does not
// expose ec.dc.* params) STATUS = -2.
//
// Mapping notes: the endpoint exposes a single simulated/real master
// link, so sNetId selects nothing beyond "a master is targeted" — a
// nonempty net id enables sync, an empty one disables it.  The
// documented 10-cycle internal/external diff check is reduced to the
// per-call |time_diff_ns| <= nSyncWindow comparison the service
// reports.
//
// SPDX-License-Identifier: Apache-2.0 OR MPL-2.0

// ---- FB_EcExtSyncExtTimes: enable/disable DC sync -----------------
// Nonempty sNetId enables ec.dc.sync_enabled and polls until the
// link reports it; bTS1Done then stays set while enabled.  Empty
// sNetId disables sync.  bError/nErrorId latch the last nonzero
// service status.

FUNCTION_BLOCK FB_EcExtSyncExtTimes
VAR_INPUT
    sNetId : STRING[22];   // T_AMSNetId
END_VAR
VAR_OUTPUT
    bTS1Done : BOOL;
    bError   : BOOL;
    nErrorId : UDINT;
END_VAR
VAR
    ch    : FB_EcSync;
    prev  : BOOL;   // previous "target present" level
    armed : BOOL;
END_VAR
    bError := FALSE;
    nErrorId := 0;

    ch.OP := 1;
    ch();
    IF ch.STATUS < 0 THEN
        bError := TRUE;
        nErrorId := ch.ERRID;
    END_IF;

    IF LEN(sNetId) > 0 AND NOT prev THEN
        ch.OP := 2;
        ch.ENABLE := 1;
        ch();
        IF ch.STATUS < 0 THEN
            bError := TRUE;
            nErrorId := ch.ERRID;
        ELSE
            armed := TRUE;
        END_IF;
        ch.OP := 1;
    ELSIF LEN(sNetId) = 0 AND prev THEN
        ch.OP := 2;
        ch.ENABLE := 0;
        ch();
        IF ch.STATUS < 0 THEN
            bError := TRUE;
            nErrorId := ch.ERRID;
        END_IF;
        ch.OP := 1;
        bTS1Done := FALSE;
        armed := FALSE;
    END_IF;

    bTS1Done := armed AND ch.CONNECTED <> 0 AND ch.SYNCEN <> 0;
    prev := LEN(sNetId) > 0;
END_FUNCTION_BLOCK

// ---- FB_EcExtSyncIsSynchronized: windowed sync check ---------------
// Polls the status op once per call.  bNotConnected is set when the
// service is unavailable or the master link is down; bSynchronized
// is set only when connected, sync enabled, and |time_diff_ns| is
// within nSyncWindow nanoseconds.

FUNCTION_BLOCK FB_EcExtSyncIsSynchronized
VAR_INPUT
    nSyncWindow : UDINT;   // nanoseconds
END_VAR
VAR_OUTPUT
    bSynchronized : BOOL;
    bNotConnected : BOOL;
    bError         : BOOL;
    nErrorId       : UDINT;
END_VAR
VAR
    ch : FB_EcSync;
    d  : LREAL;
    w  : LREAL;
END_VAR
    bError := FALSE;
    nErrorId := 0;

    ch.OP := 1;
    ch();
    IF ch.STATUS < 0 THEN
        bError := TRUE;
        nErrorId := ch.ERRID;
    END_IF;

    bSynchronized := FALSE;
    bNotConnected := FALSE;
    IF ch.STATUS < 0 OR ch.CONNECTED = 0 THEN
        bNotConnected := TRUE;
    ELSIF ch.SYNCEN <> 0 THEN
        d := ch.DIFFNS;
        IF d < 0.0 THEN d := -d; END_IF;
        w := nSyncWindow;
        IF d <= w THEN
            bSynchronized := TRUE;
        END_IF;
    END_IF;
END_FUNCTION_BLOCK

(* ---- tc3_eventlog.st ---- *)
// Tc3_EventLogger -> FB_TcEvent / FB_TcMessage / FB_TcAlarm over
// the tplc-eventlog bounded journal (128 entries, deterministic).
// Documented reductions vs the 146-entry catalogue:
//   - METHOD calls are edge-triggered command inputs (nCmd):
//     FB_TcEvent: 1=Create+Send 2=Clear 3=Confirm.
//   - Event classes are UDINT ids (no GUID type in this ST).
//   - Text args are passed raw (nArgs pack) — no .tmx resource
//     lookup or language switching; text is a literal STRING.
//   - Async text-request / remote-logger families are modelled
//     synchronously: FB_TcEventQuery covers journal reads and
//     FB_TcEventBase.RequestEventText/ClassName copy descriptor
//     fields (no .tmx resource lookup, no ADS notifications —
//     FB_TcRemoteEventLogger stays a documented gap).
//   - nErrId carries tplc-eventlog service codes.

// ---- FB_TcEvent: create/raise/clear/confirm one event ----
FUNCTION_BLOCK FB_TcEvent
VAR_INPUT
    nCmd : UDINT;               // 0 none, 1 raise, 2 clear, 3 confirm
    nEventClass : UDINT;
    nEventId : UDINT;
    nSeverity : UDINT;          // 0 verbose..4 critical
    sText : STRING[80];
    nArgs : UDINT;
END_VAR
VAR_OUTPUT
    hEvent : UDINT;             // journal id, 0 = none
    nState : UDINT;             // 1 raised 2 cleared 3 confirmed
    bDone : BOOL;
    bBusy : BOOL;
    bError : BOOL;
    nErrId : UDINT;
END_VAR
VAR
    ev : FB_EventLog;
    prev : UDINT;
END_VAR
    bDone := FALSE; bError := FALSE; nErrId := 0; bBusy := FALSE;
    IF nCmd <> 0 AND prev = 0 THEN
        bBusy := TRUE;
        ev.ID := hEvent;
        IF nCmd = 1 THEN
            ev.OP := 1; ev.ECLASS := nEventClass;
            ev.EVTID := nEventId; ev.SEV := nSeverity;
            ev.ARGS := nArgs;
            ev.TEXT := sText;
        ELSIF nCmd = 2 THEN
            ev.OP := 2;
        ELSIF nCmd = 3 THEN
            ev.OP := 3;
        END_IF;
        ev();
        IF ev.STATUS = 0 THEN
            bDone := TRUE; bBusy := FALSE;
            IF nCmd = 1 THEN
                hEvent := ev.ID; nState := 1;
            ELSIF nCmd = 2 THEN
                nState := 2;
            ELSE
                nState := 3; hEvent := 0;
            END_IF;
        ELSE
            bError := TRUE; nErrId := ev.ERRID;
        END_IF;
    END_IF;
    prev := nCmd;
END_FUNCTION_BLOCK

// ---- FB_TcMessage: INFO-severity event (send/reset) ----
FUNCTION_BLOCK FB_TcMessage
VAR_INPUT
    nCmd : UDINT;               // 1 send, 3 confirm+forget
    nEventClass : UDINT;
    nEventId : UDINT;
    sText : STRING[80];
    nArgs : UDINT;
END_VAR
VAR_OUTPUT
    hEvent : UDINT;
    bDone : BOOL;
    bError : BOOL;
    nErrId : UDINT;
END_VAR
VAR
    ev : FB_TcEvent;
END_VAR
    bDone := FALSE; bError := FALSE; nErrId := 0;
    ev.nCmd := nCmd;
    ev.nEventClass := nEventClass;
    ev.nEventId := nEventId;
    ev.nSeverity := 1;              // INFO
    ev.sText := sText;
    ev.nArgs := nArgs;
    ev();
    hEvent := ev.hEvent;
    bDone := ev.bDone;
    bError := ev.bError;
    nErrId := ev.nErrId;
END_FUNCTION_BLOCK

// ---- FB_TcAlarm: raisable/clearable/confirmable alarm ----
FUNCTION_BLOCK FB_TcAlarm
VAR_INPUT
    nCmd : UDINT;               // 1 raise, 2 clear, 3 confirm
    nEventClass : UDINT;
    nEventId : UDINT;
    nSeverity : UDINT;          // typically WARNING/ERROR
    sText : STRING[80];
    nArgs : UDINT;
END_VAR
VAR_OUTPUT
    hEvent : UDINT;
    nState : UDINT;
    bActive : BOOL;             // raised and not confirmed
    bDone : BOOL;
    bError : BOOL;
    nErrId : UDINT;
END_VAR
VAR
    ev : FB_TcEvent;
END_VAR
    bDone := FALSE; bError := FALSE; nErrId := 0;
    ev.nCmd := nCmd;
    ev.nEventClass := nEventClass;
    ev.nEventId := nEventId;
    ev.nSeverity := nSeverity;
    ev.sText := sText;
    ev.nArgs := nArgs;
    ev();
    hEvent := ev.hEvent;
    nState := ev.nState;
    bDone := ev.bDone;
    bError := ev.bError;
    nErrId := ev.nErrId;
    bActive := ev.nState = 1 OR ev.nState = 2;
END_FUNCTION_BLOCK

// ---- FB_TcEventQuery: synchronous journal read + stats ----
FUNCTION_BLOCK FB_TcEventQuery
VAR_INPUT
    nCmd : UDINT;               // 4 query, 5 stats
    nId : UDINT;
END_VAR
VAR_OUTPUT
    nState : UDINT;
    nSeverity : UDINT;
    nEventClass : UDINT;
    nEventId : UDINT;
    sText : STRING[80];
    nLive : UDINT;
    nRaised : UDINT;
    nCleared : UDINT;
    nConfirmed : UDINT;
    nDropped : UDINT;
    tRaised : ULINT;            // realtime ns at raise (0 = n/a)
    tCleared : ULINT;           // realtime ns at clear
    tConfirmed : ULINT;         // realtime ns at confirm
    bDone : BOOL;
    bError : BOOL;
    nErrId : UDINT;
END_VAR
VAR
    ev : FB_EventLog;
    prev : UDINT;
END_VAR
    bDone := FALSE; bError := FALSE; nErrId := 0;
    IF nCmd <> 0 AND prev = 0 THEN
        IF nCmd = 4 OR nCmd = 5 THEN
            ev.OP := nCmd; ev.ID := nId;
            ev();
            IF ev.STATUS = 0 THEN
                bDone := TRUE;
                IF nCmd = 4 THEN
                    nState := ev.STATE;
                    nSeverity := ev.SEVO;
                    nEventClass := ev.CLSO;
                    nEventId := ev.EVTIDO;
                    sText := ev.TXTO;
                    tRaised := ev.TSTAMP;
                    tCleared := ev.CSTAMP;
                    tConfirmed := ev.FSTAMP;
                ELSE
                    nLive := ev.LIVE;
                    nRaised := ev.RAISED;
                    nCleared := ev.CLEARED;
                    nConfirmed := ev.CONFIRMED;
                    nDropped := ev.DROPPED;
                END_IF;
            ELSE
                bError := TRUE; nErrId := ev.ERRID;
            END_IF;
        END_IF;
    END_IF;
    prev := nCmd;
END_FUNCTION_BLOCK

// ---- helpers ----
// UDINT -> decimal text (no STRING_TO_UDINT builtin)
FUNCTION F_ElU32Str : STRING[10]
VAR_INPUT
    v : UDINT;
END_VAR
VAR
    x : UDINT;
    d : UDINT;
    s : STRING[10];
    c : STRING[1];
END_VAR
    IF v = 0 THEN
        F_ElU32Str := '0';
        RETURN;
    END_IF;
    x := v; s := '';
    WHILE x > 0 DO
        d := x MOD 10;
        CASE d OF
            0: c := '0';  1: c := '1';  2: c := '2';  3: c := '3';
            4: c := '4';  5: c := '5';  6: c := '6';  7: c := '7';
            8: c := '8';  ELSE c := '9';
        END_CASE;
        s := CONCAT(c, s);
        x := x / 10;
    END_WHILE;
    F_ElU32Str := s;
END_FUNCTION

// string equality via FIND (direct = is not usable on strings)
FUNCTION F_ElStreq : BOOL
VAR_INPUT
    a : STRING[80];
    b : STRING[80];
END_VAR
    F_ElStreq := LEN(a) = LEN(b) AND FIND(a, b) = 1;
END_FUNCTION

// ---- FB_TcEventBase: event descriptor + comparisons ----
// Descriptor fields (EventClass/EventId/Severity/Text) are public
// members set directly, mirroring the TwinCAT property surface;
// nCmd selects the METHOD-equivalent operation.
FUNCTION_BLOCK FB_TcEventBase
VAR_INPUT
    nCmd : UDINT;               // 1 EqualsTo 2 EqualsToEventClass
                                // 3 EqualsToEventEntry 4 GetJsonAttr
                                // 5 RequestEventClassName
                                // 6 RequestEventText 7 Release
    cClass : UDINT;
    cId : UDINT;
    cSev : UDINT;
    cText : STRING[80];
    cEntryId : UDINT;           // journal id for EqualsToEventEntry
    sAttr : STRING[31];         // 'class' 'id' 'severity' 'text'
END_VAR
VAR_OUTPUT
    bEqual : BOOL;
    sOut : STRING[80];
    bDone : BOOL;
    bError : BOOL;
    nErrId : UDINT;
END_VAR
VAR
    prev : UDINT;
    ev : FB_EventLog;
    // public descriptor members (TwinCAT ipEventClass etc.)
    EventClass : UDINT;
    EventId : UDINT;
    Severity : UDINT;
    Text : STRING[80];
END_VAR
    bDone := FALSE; bError := FALSE; nErrId := 0; bEqual := FALSE;
    sOut := '';
    IF nCmd <> 0 AND prev = 0 THEN
        IF nCmd = 7 THEN
            EventClass := 0; EventId := 0; Severity := 0; Text := '';
            bDone := TRUE;
        ELSIF nCmd = 1 THEN
            bEqual := EventClass = cClass AND EventId = cId
                      AND Severity = cSev AND F_ElStreq(Text, cText);
            bDone := TRUE;
        ELSIF nCmd = 2 THEN
            bEqual := EventClass = cClass;
            bDone := TRUE;
        ELSIF nCmd = 3 THEN
            ev.OP := 4; ev.ID := cEntryId; ev();
            IF ev.STATUS = 0 THEN
                bEqual := EventClass = ev.CLSO AND EventId = ev.EVTIDO
                          AND Severity = ev.SEVO
                          AND F_ElStreq(Text, ev.TXTO);
            ELSE
                bError := TRUE; nErrId := ev.ERRID;
            END_IF;
            bDone := TRUE;
        ELSIF nCmd = 4 THEN
            IF F_ElStreq(sAttr, 'class') THEN
                sOut := F_ElU32Str(EventClass);
            ELSIF F_ElStreq(sAttr, 'id') THEN
                sOut := F_ElU32Str(EventId);
            ELSIF F_ElStreq(sAttr, 'severity') THEN
                sOut := F_ElU32Str(Severity);
            ELSIF F_ElStreq(sAttr, 'text') THEN
                sOut := Text;
            ELSE
                bError := TRUE; nErrId := 6;
            END_IF;
            bDone := TRUE;
        ELSIF nCmd = 5 THEN
            // no class-name table: the class id is the name
            sOut := F_ElU32Str(EventClass);
            bDone := TRUE;
        ELSIF nCmd = 6 THEN
            sOut := Text;
            bDone := TRUE;
        END_IF;
    END_IF;
    prev := nCmd;
END_FUNCTION_BLOCK

// ---- FB_TcArguments: typed argument list (I_TcArguments) ----
// METHODS Add* become commands; values are kept in fixed arrays
// (8 slots).  IsEmpty/nCount are live outputs.
FUNCTION_BLOCK FB_TcArguments
VAR_INPUT
    nCmd : UDINT;               // 1 AddInt 2 AddReal 3 AddString
                                // 4 AddBool 5 Clear
    nInt : DINT;
    fReal : LREAL;
    sArg : STRING[31];
    bArg : BOOL;
END_VAR
VAR_OUTPUT
    nCount : UDINT;
    bEmpty : BOOL;
    bDone : BOOL;
    bError : BOOL;
    nErrId : UDINT;
END_VAR
VAR
    prev : UDINT;
    cnt : UDINT;
    kd : ARRAY[0..7] OF INT;    // 1 int 2 real 3 string 4 bool
    iv : ARRAY[0..7] OF DINT;
    fv : ARRAY[0..7] OF LREAL;
    sv : ARRAY[0..7] OF STRING[31];
    bv : ARRAY[0..7] OF BOOL;
END_VAR
    bDone := FALSE; bError := FALSE; nErrId := 0;
    nCount := cnt; bEmpty := cnt = 0;
    IF nCmd <> 0 AND prev = 0 THEN
        IF nCmd = 5 THEN
            cnt := 0; bDone := TRUE;
        ELSE
            IF cnt >= 8 THEN
                bError := TRUE; nErrId := 3;
            ELSE
                IF nCmd = 1 THEN
                    kd[cnt] := 1; iv[cnt] := nInt;
                ELSIF nCmd = 2 THEN
                    kd[cnt] := 2; fv[cnt] := fReal;
                ELSIF nCmd = 3 THEN
                    kd[cnt] := 3; sv[cnt] := sArg;
                ELSIF nCmd = 4 THEN
                    kd[cnt] := 4; bv[cnt] := bArg;
                ELSE
                    bError := TRUE; nErrId := 1;
                END_IF;
                IF NOT bError THEN
                    cnt := cnt + 1; bDone := TRUE;
                END_IF;
            END_IF;
        END_IF;
    END_IF;
    prev := nCmd;
END_FUNCTION_BLOCK

// ---- FB_TcSourceInfo: source-name descriptor ----
// Name/Extended are public members; nCmd mirrors Clear /
// ExtendName / ResetToDefault.
FUNCTION_BLOCK FB_TcSourceInfo
VAR_INPUT
    nCmd : UDINT;               // 1 ExtendName 2 ResetToDefault
                                // 3 Clear
END_VAR
VAR_OUTPUT
    bDone : BOOL;
    bError : BOOL;
    nErrId : UDINT;
END_VAR
VAR
    prev : UDINT;
    Name : STRING[31];
    Extended : BOOL;
END_VAR
    bDone := FALSE; bError := FALSE; nErrId := 0;
    IF nCmd <> 0 AND prev = 0 THEN
        IF nCmd = 1 THEN
            Extended := TRUE; bDone := TRUE;
        ELSIF nCmd = 2 THEN
            Extended := FALSE; bDone := TRUE;
        ELSIF nCmd = 3 THEN
            Name := ''; Extended := FALSE; bDone := TRUE;
        END_IF;
    END_IF;
    prev := nCmd;
END_FUNCTION_BLOCK

// ---- FB_TcCauseRemedy: cause/remedy text carrier ----
// Id/Cause/Remedy are public members; nCmd 1 loads them from the
// inputs (TwinCAT GetCause/GetId/GetRemedy read members directly),
// nCmd 2 releases.
FUNCTION_BLOCK FB_TcCauseRemedy
VAR_INPUT
    nCmd : UDINT;               // 1 Load 2 Release
    nId : UDINT;
    sCause : STRING[31];
    sRemedy : STRING[31];
END_VAR
VAR_OUTPUT
    bDone : BOOL;
    bError : BOOL;
    nErrId : UDINT;
END_VAR
VAR
    prev : UDINT;
    Id : UDINT;
    Cause : STRING[31];
    Remedy : STRING[31];
END_VAR
    bDone := FALSE; bError := FALSE; nErrId := 0;
    IF nCmd <> 0 AND prev = 0 THEN
        IF nCmd = 1 THEN
            Id := nId; Cause := sCause; Remedy := sRemedy;
            bDone := TRUE;
        ELSIF nCmd = 2 THEN
            Id := 0; Cause := ''; Remedy := '';
            bDone := TRUE;
        END_IF;
    END_IF;
    prev := nCmd;
END_FUNCTION_BLOCK

// ---- FB_TcDetail: name/text/comment carrier (same shape) ----
FUNCTION_BLOCK FB_TcDetail
VAR_INPUT
    nCmd : UDINT;               // 1 Load 2 Release
    sName : STRING[31];
    sText : STRING[31];
    sComment : STRING[31];
END_VAR
VAR_OUTPUT
    bDone : BOOL;
    bError : BOOL;
    nErrId : UDINT;
END_VAR
VAR
    prev : UDINT;
    Name : STRING[31];
    Text : STRING[31];
    Comment : STRING[31];
END_VAR
    bDone := FALSE; bError := FALSE; nErrId := 0;
    IF nCmd <> 0 AND prev = 0 THEN
        IF nCmd = 1 THEN
            Name := sName; Text := sText; Comment := sComment;
            bDone := TRUE;
        ELSIF nCmd = 2 THEN
            Name := ''; Text := ''; Comment := '';
            bDone := TRUE;
        END_IF;
    END_IF;
    prev := nCmd;
END_FUNCTION_BLOCK

// ---- FB_TcEventLogger: aggregate logger surface ----
// nCmd: 1 SendMessage 2 ClearAlarms(filter) 3 ClearAllAlarms
//       4 ClearLoggedEvents 5 ConfirmAlarms(filter)
//       6 ConfirmAllAlarms 7 IsAlarmRaised(filter)
//       8 GetAlarm(filter) 9 ExportLoggedEvents
// "Alarm" = severity >= WARNING (2); filter wildcards are 0.
FUNCTION_BLOCK FB_TcEventLogger
VAR_INPUT
    nCmd : UDINT;
    nEventClass : UDINT;
    nEventId : UDINT;
    nSeverity : UDINT;
    sText : STRING[80];
    nArgs : UDINT;
    nFilterClass : UDINT;       // 0 = any class
    nFilterEid : UDINT;         // 0 = any event id
END_VAR
VAR_OUTPUT
    hEvent : UDINT;
    bFound : BOOL;
    nCount : UDINT;
    nState : UDINT;
    nSevOut : UDINT;
    nClassOut : UDINT;
    nEidOut : UDINT;
    sTextOut : STRING[80];
    sExport : STRING[255];
    bTruncated : BOOL;
    bDone : BOOL;
    bBusy : BOOL;
    bError : BOOL;
    nErrId : UDINT;
END_VAR
VAR
    ev : FB_EventLog;
    msg : FB_TcMessage;
    prev : UDINT;
    i : UDINT;
    hit : BOOL;
    filt : BOOL;
    piece : STRING[255];
END_VAR
    bDone := FALSE; bBusy := FALSE; bError := FALSE; nErrId := 0;
    bFound := FALSE; nCount := 0; bTruncated := FALSE; sExport := '';
    IF nCmd <> 0 AND prev = 0 THEN
        IF nCmd = 1 THEN
            msg.nCmd := 1;
            msg.nEventClass := nEventClass;
            msg.nEventId := nEventId;
            msg.sText := sText;
            msg.nArgs := nArgs;
            msg();
            IF msg.bDone THEN
                hEvent := msg.hEvent; bDone := TRUE;
            ELSE
                bError := TRUE; nErrId := msg.nErrId;
            END_IF;
        ELSE
            FOR i := 1 TO 128 DO
                ev.OP := 4; ev.ID := i; ev();
                IF ev.STATUS = 0 THEN
                    filt := nCmd = 3
                            OR ((nFilterClass = 0 OR ev.CLSO = nFilterClass)
                                AND (nFilterEid = 0
                                     OR ev.EVTIDO = nFilterEid));
                    hit := filt AND ev.SEVO >= 2;
                    IF nCmd = 9 THEN
                        // export every live entry as a CSV row
                        piece := CONCAT(F_ElU32Str(i), ';');
                        piece := CONCAT(piece, F_ElU32Str(ev.CLSO));
                        piece := CONCAT(piece, ';');
                        piece := CONCAT(piece, F_ElU32Str(ev.EVTIDO));
                        piece := CONCAT(piece, ';');
                        piece := CONCAT(piece, F_ElU32Str(ev.SEVO));
                        piece := CONCAT(piece, ';');
                        piece := CONCAT(piece, F_ElU32Str(ev.STATE));
                        piece := CONCAT(piece, ';');
                        piece := CONCAT(piece, ev.TXTO);
                        piece := CONCAT(piece, '|');
                        IF LEN(sExport) + LEN(piece) < 250 THEN
                            sExport := CONCAT(sExport, piece);
                        ELSE
                            bTruncated := TRUE;
                        END_IF;
                    ELSIF hit AND ev.STATE <> 3 THEN
                        // candidate alarm entry
                        // (nCmd 6 is handled by the post-loop pass)
                        IF (nCmd = 2 AND ev.STATE = 1) OR nCmd = 5
                           OR nCmd = 3 THEN
                            IF nCmd = 5 THEN
                                ev.OP := 3; ev.ID := i; ev();
                            ELSE
                                ev.OP := 2; ev.ID := i; ev();
                            END_IF;
                            IF ev.STATUS = 0 THEN nCount := nCount + 1; END_IF;
                        END_IF;
                        IF NOT bFound
                           AND (nCmd = 7 OR nCmd = 8) THEN
                            bFound := TRUE;
                            nState := ev.STATE;
                            nSevOut := ev.SEVO;
                            nClassOut := ev.CLSO;
                            nEidOut := ev.EVTIDO;
                            sTextOut := ev.TXTO;
                        END_IF;
                    END_IF;
                END_IF;
            END_FOR;
            IF nCmd = 4 THEN
                // ClearLoggedEvents: confirm every non-terminal entry
                FOR i := 1 TO 128 DO
                    ev.OP := 4; ev.ID := i; ev();
                    IF ev.STATUS = 0 AND ev.STATE <> 3 THEN
                        ev.OP := 3; ev.ID := i; ev();
                        IF ev.STATUS = 0 THEN nCount := nCount + 1; END_IF;
                    END_IF;
                END_FOR;
            END_IF;
            IF nCmd = 6 THEN
                // ConfirmAllAlarms ignores the filter
                FOR i := 1 TO 128 DO
                    ev.OP := 4; ev.ID := i; ev();
                    IF ev.STATUS = 0 AND ev.STATE <> 3 AND ev.SEVO >= 2 THEN
                        ev.OP := 3; ev.ID := i; ev();
                        IF ev.STATUS = 0 THEN nCount := nCount + 1; END_IF;
                    END_IF;
                END_FOR;
            END_IF;
            bDone := TRUE;
        END_IF;
    END_IF;
    prev := nCmd;
END_FUNCTION_BLOCK

(* ---- tc3_ftp.st ---- *)
// Tc3_FTP + Tc2_FTP -> FTP client wrappers (RFC 959, PASV data mode).
// TwinCAT's FB_FtpConnection/FB_FtpExplorer/FB_FtpTransfer objects
// and the Tc2_FTP FB_* blocks map onto the poll-driven service
// model used by the other compat libraries: FB_FtpConn holds the
// control session, FB_FtpCmd runs one control command per EXEC
// edge, FB_FtpXfer runs one RETR/STOR/LIST data transfer.
// Differences from the TwinCAT FBs, documented in
// docs/plc/compat/README.md:
//   - No FTP profile objects (AddProfile/GetProfile), no AMS/ADS
//     routing, no I_TcMessage/EventLogger/HRESULT surfaces.
//     Credentials are plain STRING inputs per connection.
//   - Passive (PASV) data connections only: no PORT/active mode,
//     no EPSV, no FTPS/TLS, no SFTP/SSH, no REST resume, no
//     MLSD/MLST, IPv4 dotted-quad hosts only (no DNS —
//     FB_FTP_HostResolve is a documented gap).
//   - Rename/move is RNFR+RNTO (works for files and directories
//     on most servers); true server-side rename semantics depend
//     on the FTP server.
//   - Downloads stream 512-byte chunks per scan (BUF + CHUNK +
//     TOTAL); uploads take UP_DATA[0..UP_LEN) once per EXEC.
//   - nStatus: conn 0=pending 1=ready 2=error; cmd 0=pending
//     1=ok(2xx) 2=fail(4xx/5xx) 3=timeout 4=error 5=badresp;
//     xfer adds 6=more-data-expected while streaming.
// Sources: docs/plc/plan/21-twincat-libraries.md (Tc2_FTP,
// Tc3_FTP).

// Open/poll/close an FTP control connection — covers
// FB_FtpConnection.Connect/Disconnect and FB_FTP_Open/
// FB_FTP_OpenEX/FB_FTP_Close/FB_FTP_Info.
FUNCTION_BLOCK FB_FTP_Connect
VAR_INPUT
    sHost : STRING[15];          // dotted-quad PLC IPv4
    nPort : UDINT := 0;          // 0 = 21
    sUser : STRING[31] := 'anonymous';
    sPass : STRING[31] := '';
    bExecute : BOOL;             // rising edge = (re)connect
    bClose : BOOL;               // rising edge = disconnect
    tTimeout : TIME := T#10S;
END_VAR
VAR_OUTPUT
    nConnHandle : UDINT;         // 0 = no live session
    bBusy : BOOL;
    bDone : BOOL;
    bError : BOOL;
    nStatus : DINT;              // 0=pending 1=ready 2=error
    nErrId : UDINT;
END_VAR
VAR
    conn : FB_FtpConn;
END_VAR
    conn.HOST := sHost;
    conn.PORT := nPort;
    conn.USER := sUser;
    conn.PASS := sPass;
    conn.TIMEOUT := tTimeout;
    conn.CLOSE := bClose;
    conn.EXEC := bExecute;
    conn();
    nConnHandle := conn.CONN_HANDLE;
    bBusy := conn.BUSY;
    bDone := conn.DONE;
    nStatus := conn.STATUS;
    nErrId := conn.ERRID;
    bError := (conn.ERRID <> 0) OR (conn.STATUS = 2);
END_FUNCTION_BLOCK

// One FTP control command — covers the explorer operations
// (MKD/RMD/DELE/RNFR/RNTO/CWD/PWD/SIZE/TYPE/SYST/NOOP/SITE)
// and is the building block for the method wrappers below.
FUNCTION_BLOCK FB_FTP_Cmd
VAR_INPUT
    nConnHandle : UDINT;         // from FB_FTP_Connect
    sCmd : STRING[127];          // e.g. 'MKD /dir'
    bExecute : BOOL;
    tTimeout : TIME := T#5S;
END_VAR
VAR_OUTPUT
    bBusy : BOOL;
    bDone : BOOL;
    bError : BOOL;
    nStatus : DINT;              // 0=pending 1=ok 2=fail 3=timeout 4=error 5=badresp
    nRespCode : UDINT;           // final 3-digit FTP reply code
    nErrId : UDINT;
    sText : STRING[127];         // reply text (last line)
END_VAR
VAR
    c : FB_FtpCmd;
END_VAR
    c.CONN_HANDLE := nConnHandle;
    c.CMD := sCmd;
    c.TIMEOUT := tTimeout;
    c.EXEC := bExecute;
    c();
    bBusy := c.BUSY;
    bDone := c.DONE;
    nStatus := c.STATUS;
    nRespCode := c.RESP_CODE;
    nErrId := c.ERRID;
    sText := c.TEXT;
    bError := (c.ERRID <> 0) OR (c.STATUS >= 2);
END_FUNCTION_BLOCK

// Download a remote file (RETR) — covers
// FB_FtpTransfer.Download and FB_FTP_FileDownload(FileDownloadEx).
// DATA receives up to 512 bytes per BUSY scan; append chunks at
// nChunk until nStatus leaves 0/6.
FUNCTION_BLOCK FB_FTP_Download
VAR_INPUT
    nConnHandle : UDINT;
    sRemotePath : STRING[127];
    bExecute : BOOL;
    tTimeout : TIME := T#30S;
END_VAR
VAR_OUTPUT
    bBusy : BOOL;
    bDone : BOOL;
    bError : BOOL;
    nStatus : DINT;              // 0=pending 6=more 1=ok 2..5=fail
    nRespCode : UDINT;
    nTotal : UDINT;              // bytes received so far
    nChunk : UDINT;              // bytes in DATA this scan
    DATA : ARRAY[0..511] OF BYTE; // latest chunk
END_VAR
VAR
    x : FB_FtpXfer;
END_VAR
    x.CONN_HANDLE := nConnHandle;
    x.OP := 0;
    x.PATH := sRemotePath;
    x.TIMEOUT := tTimeout;
    x.EXEC := bExecute;
    x();
    bBusy := x.BUSY;
    bDone := x.DONE;
    nStatus := x.STATUS;
    nRespCode := x.RESP_CODE;
    nTotal := x.TOTAL;
    nChunk := x.CHUNK;
    DATA := x.BUF;
    bError := (x.ERRID <> 0) OR ((x.STATUS >= 1) AND (x.STATUS <= 5));
END_FUNCTION_BLOCK

// Upload a local file (STOR) — covers FB_FtpTransfer.Upload and
// FB_FTP_FileUpload(FileUploadEx). DATA holds the bytes to send
// (nLen valid, <= 512 per transfer).
FUNCTION_BLOCK FB_FTP_Upload
VAR_INPUT
    nConnHandle : UDINT;
    sRemotePath : STRING[127];
    nLen : UDINT;                // bytes in DATA, <= 512
    DATA : ARRAY[0..511] OF BYTE;
    bExecute : BOOL;
    tTimeout : TIME := T#30S;
END_VAR
VAR_OUTPUT
    bBusy : BOOL;
    bDone : BOOL;
    bError : BOOL;
    nStatus : DINT;
    nRespCode : UDINT;
    nTotal : UDINT;              // bytes accepted/sent so far
END_VAR
VAR
    x : FB_FtpXfer;
    i : UDINT;
END_VAR
    x.CONN_HANDLE := nConnHandle;
    x.OP := 1;
    x.PATH := sRemotePath;
    x.TIMEOUT := tTimeout;
    x.UP_LEN := nLen;
    FOR i := 0 TO 511 DO
        x.UP_DATA[i] := DATA[i];
    END_FOR;
    x.EXEC := bExecute;
    x();
    bBusy := x.BUSY;
    bDone := x.DONE;
    nStatus := x.STATUS;
    nRespCode := x.RESP_CODE;
    nTotal := x.TOTAL;
    bError := (x.ERRID <> 0) OR ((x.STATUS >= 1) AND (x.STATUS <= 5));
END_FUNCTION_BLOCK

// List a remote directory (LIST/NLST) — covers
// FB_FTP_FileList(FileListEx) and the explorer listing path.
// Same chunked download semantics as FB_FTP_Download.
FUNCTION_BLOCK FB_FTP_List
VAR_INPUT
    nConnHandle : UDINT;
    sRemotePath : STRING[127];   // '' = current directory
    bExecute : BOOL;
    tTimeout : TIME := T#30S;
END_VAR
VAR_OUTPUT
    bBusy : BOOL;
    bDone : BOOL;
    bError : BOOL;
    nStatus : DINT;
    nRespCode : UDINT;
    nTotal : UDINT;
    nChunk : UDINT;
    DATA : ARRAY[0..511] OF BYTE; // latest listing chunk
END_VAR
VAR
    x : FB_FtpXfer;
END_VAR
    x.CONN_HANDLE := nConnHandle;
    x.OP := 2;
    x.PATH := sRemotePath;
    x.TIMEOUT := tTimeout;
    x.EXEC := bExecute;
    x();
    bBusy := x.BUSY;
    bDone := x.DONE;
    nStatus := x.STATUS;
    nRespCode := x.RESP_CODE;
    nTotal := x.TOTAL;
    nChunk := x.CHUNK;
    DATA := x.BUF;
    bError := (x.ERRID <> 0) OR ((x.STATUS >= 1) AND (x.STATUS <= 5));
END_FUNCTION_BLOCK

// Create a remote directory — covers FB_FtpExplorer.DirCreate
// and FB_FTP_DirCreate.
FUNCTION_BLOCK FB_FTP_MkDir
VAR_INPUT
    nConnHandle : UDINT;
    sPath : STRING[127];
    bExecute : BOOL;
    tTimeout : TIME := T#5S;
END_VAR
VAR_OUTPUT
    bBusy : BOOL;
    bDone : BOOL;
    bError : BOOL;
    nStatus : DINT;
    nRespCode : UDINT;
    nErrId : UDINT;
END_VAR
VAR
    c : FB_FTP_Cmd;
    sCmd : STRING[127];
END_VAR
    sCmd := CONCAT('MKD ', sPath);
    c.nConnHandle := nConnHandle;
    c.sCmd := sCmd;
    c.tTimeout := tTimeout;
    c.bExecute := bExecute;
    c();
    bBusy := c.bBusy;
    bDone := c.bDone;
    nStatus := c.nStatus;
    nRespCode := c.nRespCode;
    nErrId := c.nErrId;
    bError := c.bError;
END_FUNCTION_BLOCK

// Remove an empty remote directory — covers
// FB_FtpExplorer.DirRemove and FB_FTP_DirRemove.
FUNCTION_BLOCK FB_FTP_RemoveDir
VAR_INPUT
    nConnHandle : UDINT;
    sPath : STRING[127];
    bExecute : BOOL;
    tTimeout : TIME := T#5S;
END_VAR
VAR_OUTPUT
    bBusy : BOOL;
    bDone : BOOL;
    bError : BOOL;
    nStatus : DINT;
    nRespCode : UDINT;
    nErrId : UDINT;
END_VAR
VAR
    c : FB_FTP_Cmd;
    sCmd : STRING[127];
END_VAR
    sCmd := CONCAT('RMD ', sPath);
    c.nConnHandle := nConnHandle;
    c.sCmd := sCmd;
    c.tTimeout := tTimeout;
    c.bExecute := bExecute;
    c();
    bBusy := c.bBusy;
    bDone := c.bDone;
    nStatus := c.nStatus;
    nRespCode := c.nRespCode;
    nErrId := c.nErrId;
    bError := c.bError;
END_FUNCTION_BLOCK

// Delete a remote file — covers FB_FtpExplorer.FileRemove
// and FB_FTP_FileRemove.
FUNCTION_BLOCK FB_FTP_DeleteFile
VAR_INPUT
    nConnHandle : UDINT;
    sPath : STRING[127];
    bExecute : BOOL;
    tTimeout : TIME := T#5S;
END_VAR
VAR_OUTPUT
    bBusy : BOOL;
    bDone : BOOL;
    bError : BOOL;
    nStatus : DINT;
    nRespCode : UDINT;
    nErrId : UDINT;
END_VAR
VAR
    c : FB_FTP_Cmd;
    sCmd : STRING[127];
END_VAR
    sCmd := CONCAT('DELE ', sPath);
    c.nConnHandle := nConnHandle;
    c.sCmd := sCmd;
    c.tTimeout := tTimeout;
    c.bExecute := bExecute;
    c();
    bBusy := c.bBusy;
    bDone := c.bDone;
    nStatus := c.nStatus;
    nRespCode := c.nRespCode;
    nErrId := c.nErrId;
    bError := c.bError;
END_FUNCTION_BLOCK

// Check remote file existence — covers
// FB_FtpExplorer.FileExists and FB_FTP_FileExist. Issues SIZE;
// 213 = exists, 550 = not found.
FUNCTION_BLOCK FB_FTP_FileExists
VAR_INPUT
    nConnHandle : UDINT;
    sPath : STRING[127];
    bExecute : BOOL;
    tTimeout : TIME := T#5S;
END_VAR
VAR_OUTPUT
    bBusy : BOOL;
    bDone : BOOL;
    bError : BOOL;
    bExists : BOOL;
    nStatus : DINT;
    nRespCode : UDINT;
    nErrId : UDINT;
END_VAR
VAR
    c : FB_FTP_Cmd;
    sCmd : STRING[127];
END_VAR
    sCmd := CONCAT('SIZE ', sPath);
    c.nConnHandle := nConnHandle;
    c.sCmd := sCmd;
    c.tTimeout := tTimeout;
    c.bExecute := bExecute;
    c();
    bBusy := c.bBusy;
    bDone := c.bDone;
    nStatus := c.nStatus;
    nRespCode := c.nRespCode;
    nErrId := c.nErrId;
    bExists := (c.nRespCode = 213);
    bError := c.bError AND (c.nStatus <> 2);
END_FUNCTION_BLOCK

// Check remote directory existence — covers
// FB_FtpExplorer.DirExists. Issues a LIST on the path; a
// completed transfer means the directory is listable (exists).
// No working-directory side effects.
FUNCTION_BLOCK FB_FTP_DirExists
VAR_INPUT
    nConnHandle : UDINT;
    sPath : STRING[127];
    bExecute : BOOL;
    tTimeout : TIME := T#10S;
END_VAR
VAR_OUTPUT
    bBusy : BOOL;
    bDone : BOOL;
    bError : BOOL;
    bExists : BOOL;
    nStatus : DINT;
    nRespCode : UDINT;
END_VAR
VAR
    x : FB_FtpXfer;
    sink : ARRAY[0..511] OF BYTE;
END_VAR
    x.CONN_HANDLE := nConnHandle;
    x.OP := 2;
    x.PATH := sPath;
    x.TIMEOUT := tTimeout;
    x.EXEC := bExecute;
    x();
    sink := x.BUF;
    bBusy := x.BUSY;
    bDone := x.DONE;
    nStatus := x.STATUS;
    nRespCode := x.RESP_CODE;
    bExists := (x.STATUS = 1);
    bError := (x.ERRID <> 0) OR ((x.STATUS >= 2) AND (x.STATUS <= 5));
END_FUNCTION_BLOCK

// Rename/move a remote file or directory — covers
// FB_FtpExplorer.FileRename/FileMove/DirRename/DirMove and
// FB_FTP_FileRename. Issues RNFR <old> then RNTO <new> on the
// same connection; success requires 350 then 250/2xx.
FUNCTION_BLOCK FB_FTP_Rename
VAR_INPUT
    nConnHandle : UDINT;
    sOldPath : STRING[127];
    sNewPath : STRING[127];
    bExecute : BOOL;
    tTimeout : TIME := T#10S;
END_VAR
VAR_OUTPUT
    bBusy : BOOL;
    bDone : BOOL;
    bError : BOOL;
    nStatus : DINT;              // 0=pending 1=ok 2=fail 3=timeout 4=error 5=badresp
    nRespCode : UDINT;           // final reply code (RNTO)
    nErrId : UDINT;
END_VAR
VAR
    rnfr : FB_FTP_Cmd;
    rnto : FB_FTP_Cmd;
    sCmd1 : STRING[127];
    sCmd2 : STRING[127];
    step : UDINT := 0;           // 0=RNFR 1=RNTO 2=report-fail
    prevExec : BOOL := FALSE;
END_VAR
    sCmd1 := CONCAT('RNFR ', sOldPath);
    sCmd2 := CONCAT('RNTO ', sNewPath);
    IF bExecute AND NOT prevExec THEN
        step := 0;
    END_IF;
    prevExec := bExecute;
    IF step = 0 THEN
        rnfr.nConnHandle := nConnHandle;
        rnfr.sCmd := sCmd1;
        rnfr.tTimeout := tTimeout;
        rnfr.bExecute := bExecute;
        rnfr();
        IF rnfr.bDone THEN
            IF rnfr.nRespCode = 350 THEN
                step := 1;
            ELSE
                step := 2;
            END_IF;
        END_IF;
        bBusy := rnfr.bBusy;
        bDone := FALSE;
        nStatus := rnfr.nStatus;
        nRespCode := rnfr.nRespCode;
        nErrId := rnfr.nErrId;
        bError := rnfr.bError;
    ELSIF step = 1 THEN
        rnto.nConnHandle := nConnHandle;
        rnto.sCmd := sCmd2;
        rnto.tTimeout := tTimeout;
        rnto.bExecute := TRUE;    // level-held; builtin edge-fires once
        rnto();
        IF rnto.bDone THEN
            step := 0;
        END_IF;
        bBusy := rnto.bBusy;
        bDone := rnto.bDone;
        nStatus := rnto.nStatus;
        nRespCode := rnto.nRespCode;
        nErrId := rnto.nErrId;
        bError := rnto.bError;
    ELSE
        // step 2: RNFR rejected — hold the failure visible until
        // bExecute drops, then arm for the next request
        bBusy := FALSE;
        bDone := TRUE;
        nStatus := 2;
        nRespCode := rnfr.nRespCode;
        nErrId := rnfr.nErrId;
        bError := TRUE;
        IF NOT bExecute THEN
            step := 0;
        END_IF;
    END_IF;
END_FUNCTION_BLOCK

(* ---- tc3_iec870.st ---- *)
// Tc2_IEC60870_5_10x -> IEC 60870 telecontrol wrappers (104 client
// plus pure ASDU helpers). TwinCAT's FB_IEC870_5_104Master/Slave
// and FB_IEC870_5_101/102/103TProtocol blocks are built on AMS-routed
// AO databases, PVOID buffers, POINTER TO ARRAY and generated
// server objects. TetherPLC adapts the supported surface to the
// poll-driven service model used by the other compat libraries:
// FB_Iec870Conn holds one IEC 60870-5-104 session (TCP 2404,
// STARTDT handshake), FB_Iec870Tx runs one ASDU send per EXEC edge,
// FB_Iec870Rx polls the received-ASDU queue every scan.
// Differences from the TwinCAT FBs, documented in
// docs/plc/compat/README.md:
//   - Master side only: 104 client. No 101/102/103 serial or HDLC
//     transports, no slave/server mode, no AO database, no AMS
//     NetID routing, no PVOID/HRESULT object model, no redundancy
//     groups, no file transfer, no TLS.
//   - ASDU payloads are raw info-object bytes; per-type object
//     codecs (measured-value scaling, CP24/CP56 timestamps,
//     sequence addressing expansion) stay in user code or the
//     pure helpers below.
//   - The pure helpers take flat scalar/array arguments instead
//     of TwinCAT STRUCT/STRING types: CP56Time2a is a 7-byte
//     ARRAY OF BYTE, SYSTEMTIME is six scalar outputs.
// Sources: docs/plc/plan/21-twincat-libraries.md
// (Tc2_IEC60870_5_10x), IEC 60870-5-104/-5-101, lib60870-CS104.

// Open/poll/close an IEC 60870-5-104 master connection —
// covers FB_IEC870_5_104Master and the generic
// FB_IEC870_5_10xTProtocol link layer for the TCP transport.
FUNCTION_BLOCK FB_IEC870_5_104Master
VAR_INPUT
    sHost : STRING[15];          // dotted-quad PLC IPv4
    nPort : UDINT := 0;          // 0 = 2404
    nCA_Size : UDINT := 2;       // common-address octets 1 or 2
    nCOT_Size : UDINT := 2;      // COT octets 1 or 2 (2nd = OA)
    bExecute : BOOL;             // rising edge = (re)connect
    bClose : BOOL;               // rising edge = disconnect
    tTimeout : TIME := T#5S;
    tKeepAlive : TIME := T#10S;  // TESTFR interval
END_VAR
VAR_OUTPUT
    nConnHandle : UDINT;         // 0 = no live session
    bBusy : BOOL;
    bDone : BOOL;
    bError : BOOL;
    nStatus : DINT;              // 0=pending 1=ready 2=error
    nSubState : DINT;            // 0=none 1=tcp 2=startdt 3=active
    nErrId : UDINT;
    nRxDropped : UDINT;
END_VAR
VAR
    conn : FB_Iec870Conn;
END_VAR
    conn.HOST := sHost;
    conn.PORT := nPort;
    conn.CA_SIZE := nCA_Size;
    conn.COT_SIZE := nCOT_Size;
    conn.TIMEOUT := tTimeout;
    conn.CLOSE := bClose;
    conn.EXEC := bExecute;
    conn();
    nConnHandle := conn.CONN_HANDLE;
    bBusy := conn.BUSY;
    bDone := conn.DONE;
    nStatus := conn.STATUS;
    nSubState := conn.SUBSTATE;
    nErrId := conn.ERRID;
    nRxDropped := conn.RX_DROPPED;
    bError := (conn.ERRID <> 0) OR (conn.STATUS = 2);
END_FUNCTION_BLOCK

// Send one ASDU as an I-frame — covers the master-side transmit
// path of FB_IEC870_5_104Master (cyclic/spontaneous ASDUs).
// nTypeId/nVSQ/nCOT/nCA are the raw ASDU header fields; pPayload
// carries the info-object bytes. One outstanding send per
// connection; the k-window (12 unacked I-frames) applies.
FUNCTION_BLOCK FB_IEC870_SendAsdu
VAR_INPUT
    nConnHandle : UDINT;         // from FB_IEC870_5_104Master
    nTypeId : UDINT;             // ASDU type identifier
    nVSQ : UDINT;                // raw VSQ octet (bit7 seq flag)
    nCOT : UDINT;                // encoded COT (+OA bits 8..15)
    nCA : UDINT;                 // common address
    nLen : UDINT;                // payload bytes 0..240
    pPayload : ARRAY[0..239] OF BYTE;
    bExecute : BOOL;
END_VAR
VAR_OUTPUT
    bBusy : BOOL;
    bDone : BOOL;
    bError : BOOL;
    nStatus : DINT;              // 0=pending 1=ok 2=error
    nErrId : UDINT;
END_VAR
VAR
    tx : FB_Iec870Tx;
    i : INT;
END_VAR
    tx.CONN_HANDLE := nConnHandle;
    tx.TYPE_ID := nTypeId;
    tx.VSQ := nVSQ;
    tx.COT := nCOT;
    tx.CA := nCA;
    tx.LEN := nLen;
    i := 0;
    WHILE i < 240 DO
        tx.PAYLOAD[i] := pPayload[i];
        i := i + 1;
    END_WHILE;
    tx.EXEC := bExecute;
    tx();
    bBusy := tx.BUSY;
    bDone := tx.DONE;
    nStatus := tx.STATUS;
    nErrId := tx.ERRID;
    bError := (tx.ERRID <> 0) OR (tx.STATUS = 2);
END_FUNCTION_BLOCK

// Poll one received ASDU — call every scan with the connection
// handle; bDone pulses TRUE once per delivered ASDU
// (consume-on-read). nTypeId/nVSQ/nCOT/nCA describe the raw ASDU
// header parsed per the conn COT_SIZE/CA_SIZE; pPayload holds
// the info-object bytes (nLen valid).
FUNCTION_BLOCK FB_IEC870_RecvAsdu
VAR_INPUT
    nConnHandle : UDINT;
END_VAR
VAR_OUTPUT
    bDone : BOOL;
    nTypeId : UDINT;
    nVSQ : UDINT;
    nCOT : UDINT;
    nCA : UDINT;
    nLen : UDINT;
    nIFrameSeq : UDINT;
    nErrId : UDINT;
    pPayload : ARRAY[0..239] OF BYTE;
END_VAR
VAR
    rx : FB_Iec870Rx;
    i : INT;
END_VAR
    rx.CONN_HANDLE := nConnHandle;
    rx();
    bDone := rx.DONE;
    nTypeId := rx.TYPE_ID;
    nVSQ := rx.VSQ;
    nCOT := rx.COT;
    nCA := rx.CA;
    nLen := rx.LEN;
    nIFrameSeq := rx.I_FRAME_SEQ;
    nErrId := rx.ERRID;
    IF rx.DONE THEN
        i := 0;
        WHILE i < 240 DO
            pPayload[i] := rx.PAYLOAD[i];
            i := i + 1;
        END_WHILE;
    END_IF
END_FUNCTION_BLOCK

// ------------------------------------------------------------------
// Pure helpers (TwinCAT helper FBs/functions, flat signatures)
// ------------------------------------------------------------------

// ASDU101COT_TO_STRING — cause-of-transmission type to text.
// Covers the 101/104 COT table.
FUNCTION ASDU101COT_TO_STRING : STRING[31]
VAR_INPUT
    nCOT : UDINT;                // COT type bits 0..5
END_VAR
VAR
    t : UDINT;
END_VAR
    t := nCOT AND 16#3F;
    CASE t OF
        1:  ASDU101COT_TO_STRING := 'PERIODIC';
        2:  ASDU101COT_TO_STRING := 'BACKGROUND';
        3:  ASDU101COT_TO_STRING := 'SPONTANEOUS';
        4:  ASDU101COT_TO_STRING := 'INITIALIZED';
        5:  ASDU101COT_TO_STRING := 'REQUEST';
        6:  ASDU101COT_TO_STRING := 'ACTIVATION';
        7:  ASDU101COT_TO_STRING := 'ACT_CON';
        8:  ASDU101COT_TO_STRING := 'DEACTIVATION';
        9:  ASDU101COT_TO_STRING := 'DEACT_CON';
        10: ASDU101COT_TO_STRING := 'ACT_TERMINATION';
        11: ASDU101COT_TO_STRING := 'REMOTE_TAG';
        12: ASDU101COT_TO_STRING := 'LOCAL_TAG';
        20: ASDU101COT_TO_STRING := 'UNKNOWN_TYPE';
    ELSE
        ASDU101COT_TO_STRING := 'RESERVED';
    END_CASE
END_FUNCTION

// ASDU102COT_TO_STRING — 102 (dial-up) COT table adds file-ready.
FUNCTION ASDU102COT_TO_STRING : STRING[31]
VAR_INPUT
    nCOT : UDINT;
END_VAR
VAR
    t : UDINT;
END_VAR
    t := nCOT AND 16#3F;
    CASE t OF
        1:  ASDU102COT_TO_STRING := 'PERIODIC';
        2:  ASDU102COT_TO_STRING := 'BACKGROUND';
        3:  ASDU102COT_TO_STRING := 'SPONTANEOUS';
        4:  ASDU102COT_TO_STRING := 'INITIALIZED';
        5:  ASDU102COT_TO_STRING := 'REQUEST';
        6:  ASDU102COT_TO_STRING := 'ACTIVATION';
        7:  ASDU102COT_TO_STRING := 'ACT_CON';
        8:  ASDU102COT_TO_STRING := 'DEACTIVATION';
        9:  ASDU102COT_TO_STRING := 'DEACT_CON';
        10: ASDU102COT_TO_STRING := 'ACT_TERMINATION';
        11: ASDU102COT_TO_STRING := 'REMOTE_TAG';
        12: ASDU102COT_TO_STRING := 'LOCAL_TAG';
        13: ASDU102COT_TO_STRING := 'FILE_READY';
        20: ASDU102COT_TO_STRING := 'UNKNOWN_TYPE';
    ELSE
        ASDU102COT_TO_STRING := 'RESERVED';
    END_CASE
END_FUNCTION

// ASDU103COT_TO_STRING — 103 (relay protection) COT table.
FUNCTION ASDU103COT_TO_STRING : STRING[31]
VAR_INPUT
    nCOT : UDINT;
END_VAR
VAR
    t : UDINT;
END_VAR
    t := nCOT AND 16#3F;
    CASE t OF
        1:  ASDU103COT_TO_STRING := 'PERIODIC';
        2:  ASDU103COT_TO_STRING := 'BACKGROUND';
        3:  ASDU103COT_TO_STRING := 'SPONTANEOUS';
        4:  ASDU103COT_TO_STRING := 'INITIALIZED';
        5:  ASDU103COT_TO_STRING := 'REQUEST';
        6:  ASDU103COT_TO_STRING := 'ACTIVATION';
        7:  ASDU103COT_TO_STRING := 'ACT_CON';
        8:  ASDU103COT_TO_STRING := 'DEACTIVATION';
        9:  ASDU103COT_TO_STRING := 'DEACT_CON';
        10: ASDU103COT_TO_STRING := 'ACT_TERMINATION';
        11: ASDU103COT_TO_STRING := 'REMOTE_TAG';
        12: ASDU103COT_TO_STRING := 'LOCAL_TAG';
        13: ASDU103COT_TO_STRING := 'FILE_READY';
        20: ASDU103COT_TO_STRING := 'UNKNOWN_TYPE';
    ELSE
        ASDU103COT_TO_STRING := 'RESERVED';
    END_CASE
END_FUNCTION

// ASDU101TYPEID_TO_STRING — common 101/104 ASDU type names.
FUNCTION ASDU101TYPEID_TO_STRING : STRING[31]
VAR_INPUT
    nTypeId : UDINT;
END_VAR
VAR
    t : UDINT;
END_VAR
    t := nTypeId;
    CASE t OF
        1:   ASDU101TYPEID_TO_STRING := 'M_SP_NA_1';
        2:   ASDU101TYPEID_TO_STRING := 'M_SP_TA_1';
        3:   ASDU101TYPEID_TO_STRING := 'M_DP_NA_1';
        4:   ASDU101TYPEID_TO_STRING := 'M_DP_TA_1';
        5:   ASDU101TYPEID_TO_STRING := 'M_ST_NA_1';
        6:   ASDU101TYPEID_TO_STRING := 'M_ST_TA_1';
        7:   ASDU101TYPEID_TO_STRING := 'M_BO_NA_1';
        8:   ASDU101TYPEID_TO_STRING := 'M_BO_TA_1';
        9:   ASDU101TYPEID_TO_STRING := 'M_ME_NA_1';
        10:  ASDU101TYPEID_TO_STRING := 'M_ME_TA_1';
        11:  ASDU101TYPEID_TO_STRING := 'M_ME_NB_1';
        12:  ASDU101TYPEID_TO_STRING := 'M_ME_TB_1';
        13:  ASDU101TYPEID_TO_STRING := 'M_ME_NC_1';
        14:  ASDU101TYPEID_TO_STRING := 'M_ME_TC_1';
        15:  ASDU101TYPEID_TO_STRING := 'M_IT_NA_1';
        16:  ASDU101TYPEID_TO_STRING := 'M_IT_TA_1';
        17:  ASDU101TYPEID_TO_STRING := 'M_EP_TA_1';
        18:  ASDU101TYPEID_TO_STRING := 'M_EP_TB_1';
        19:  ASDU101TYPEID_TO_STRING := 'M_EP_TC_1';
        20:  ASDU101TYPEID_TO_STRING := 'M_EP_TD_1';
        21:  ASDU101TYPEID_TO_STRING := 'M_EP_TE_1';
        30:  ASDU101TYPEID_TO_STRING := 'M_SP_TB_1';
        31:  ASDU101TYPEID_TO_STRING := 'M_DP_TB_1';
        32:  ASDU101TYPEID_TO_STRING := 'M_ST_TB_1';
        33:  ASDU101TYPEID_TO_STRING := 'M_BO_TB_1';
        34:  ASDU101TYPEID_TO_STRING := 'M_ME_TD_1';
        35:  ASDU101TYPEID_TO_STRING := 'M_ME_TE_1';
        36:  ASDU101TYPEID_TO_STRING := 'M_ME_TF_1';
        37:  ASDU101TYPEID_TO_STRING := 'M_IT_TB_1';
        38:  ASDU101TYPEID_TO_STRING := 'M_EP_TF_1';
        39:  ASDU101TYPEID_TO_STRING := 'M_EP_TG_1';
        40:  ASDU101TYPEID_TO_STRING := 'M_EP_TH_1';
        41:  ASDU101TYPEID_TO_STRING := 'M_EP_TI_1';
        42:  ASDU101TYPEID_TO_STRING := 'M_EP_TJ_1';
        43:  ASDU101TYPEID_TO_STRING := 'M_EP_TK_1';
        44:  ASDU101TYPEID_TO_STRING := 'M_EP_TL_1';
        45:  ASDU101TYPEID_TO_STRING := 'C_SC_NA_1';
        46:  ASDU101TYPEID_TO_STRING := 'C_DC_NA_1';
        47:  ASDU101TYPEID_TO_STRING := 'C_RC_NA_1';
        48:  ASDU101TYPEID_TO_STRING := 'C_SE_NA_1';
        49:  ASDU101TYPEID_TO_STRING := 'C_SE_NB_1';
        50:  ASDU101TYPEID_TO_STRING := 'C_SE_NC_1';
        51:  ASDU101TYPEID_TO_STRING := 'C_BO_NA_1';
        58:  ASDU101TYPEID_TO_STRING := 'C_SC_TA_1';
        59:  ASDU101TYPEID_TO_STRING := 'C_DC_TA_1';
        60:  ASDU101TYPEID_TO_STRING := 'C_RC_TA_1';
        61:  ASDU101TYPEID_TO_STRING := 'C_SE_TA_1';
        62:  ASDU101TYPEID_TO_STRING := 'C_SE_TB_1';
        63:  ASDU101TYPEID_TO_STRING := 'C_SE_TC_1';
        64:  ASDU101TYPEID_TO_STRING := 'C_BO_TA_1';
        70:  ASDU101TYPEID_TO_STRING := 'M_EI_NA_1';
        100: ASDU101TYPEID_TO_STRING := 'C_IC_NA_1';
        101: ASDU101TYPEID_TO_STRING := 'C_CI_NA_1';
        102: ASDU101TYPEID_TO_STRING := 'C_RD_NA_1';
        103: ASDU101TYPEID_TO_STRING := 'C_CS_NA_1';
        104: ASDU101TYPEID_TO_STRING := 'C_TS_NA_1';
        105: ASDU101TYPEID_TO_STRING := 'C_RP_NA_1';
        106: ASDU101TYPEID_TO_STRING := 'C_CD_NA_1';
        107: ASDU101TYPEID_TO_STRING := 'C_TS_TA_1';
    ELSE
        ASDU101TYPEID_TO_STRING := 'UNKNOWN';
    END_CASE
END_FUNCTION

// ASDU102TYPEID_TO_STRING / ASDU103TYPEID_TO_STRING — the 102/103
// tables share the common monitoring/command IDs with 101 plus
// file-transfer and protection-event types; the common subset
// delegates to ASDU101TYPEID_TO_STRING.
FUNCTION ASDU102TYPEID_TO_STRING : STRING[31]
VAR_INPUT
    nTypeId : UDINT;
END_VAR
VAR
    t : UDINT;
END_VAR
    t := nTypeId;
    IF (t >= 1) AND (t <= 71) THEN
        ASDU102TYPEID_TO_STRING := ASDU101TYPEID_TO_STRING(t);
    ELSIF (t >= 100) AND (t <= 107) THEN
        ASDU102TYPEID_TO_STRING := ASDU101TYPEID_TO_STRING(t);
    ELSIF (t >= 110) AND (t <= 115) THEN
        ASDU102TYPEID_TO_STRING := 'FILE_SEGMENT';
    ELSE
        ASDU102TYPEID_TO_STRING := 'UNKNOWN';
    END_IF
END_FUNCTION

FUNCTION ASDU103TYPEID_TO_STRING : STRING[31]
VAR_INPUT
    nTypeId : UDINT;
END_VAR
VAR
    t : UDINT;
END_VAR
    t := nTypeId;
    IF (t >= 1) AND (t <= 44) THEN
        ASDU103TYPEID_TO_STRING := ASDU101TYPEID_TO_STRING(t);
    ELSIF (t >= 45) AND (t <= 64) THEN
        ASDU103TYPEID_TO_STRING := ASDU101TYPEID_TO_STRING(t);
    ELSIF t = 70 THEN
        ASDU103TYPEID_TO_STRING := 'M_EI_NA_1';
    ELSIF t = 71 THEN
        ASDU103TYPEID_TO_STRING := 'M_EI_TA_1';
    ELSIF (t >= 90) AND (t <= 99) THEN
        ASDU103TYPEID_TO_STRING := 'PROTECTION_EVENT';
    ELSE
        ASDU103TYPEID_TO_STRING := 'UNKNOWN';
    END_IF
END_FUNCTION

// QOI_TO_COT — quality-of-information flags to the QDS/COT-style
// flag bits (OV=0x01, BL=0x10, SUC=0x20, IV=0x80).
FUNCTION QOI_TO_COT : UDINT
VAR_INPUT
    bIV : BOOL;                  // invalid
    bSU : BOOL;                  // substituted
    bBL : BOOL;                  // blocked
    bOV : BOOL;                  // overflow
END_VAR
VAR
    r : UDINT;
END_VAR
    r := 0;
    IF bOV THEN r := r OR 16#01; END_IF;
    IF bBL THEN r := r OR 16#10; END_IF;
    IF bSU THEN r := r OR 16#20; END_IF;
    IF bIV THEN r := r OR 16#80; END_IF;
    QOI_TO_COT := r;
END_FUNCTION

// RQT_TO_COT — request-type to COT cause for command ASDUs:
// select=activation(6), execute=activation(6),
// abort/deactivate=deactivation(8).
FUNCTION RQT_TO_COT : UDINT
VAR_INPUT
    nRqt : UDINT;
END_VAR
    IF nRqt >= 4 THEN
        RQT_TO_COT := 8;          // abort family -> deactivation
    ELSE
        RQT_TO_COT := 6;          // select/execute -> activation
    END_IF
END_FUNCTION

// CP24IOA_TO_DWORD — pack a 24-bit information object address
// (3 big-endian octets) into a DWORD for table lookups.
FUNCTION CP24IOA_TO_DWORD : UDINT
VAR_INPUT
    b0 : UDINT;                  // IOA octet 0 (MSB)
    b1 : UDINT;                  // IOA octet 1
    b2 : UDINT;                  // IOA octet 2 (LSB)
END_VAR
    CP24IOA_TO_DWORD := (b0 AND 16#FF) * 65536 +
                        (b1 AND 16#FF) * 256 +
                        (b2 AND 16#FF);
END_FUNCTION

FUNCTION DWORD_TO_CP24IOA : UDINT
VAR_INPUT
    nIOA : UDINT;                // packed 24-bit value
END_VAR
    DWORD_TO_CP24IOA := nIOA AND 16#FFFFFF;
END_FUNCTION

// CP56Time2a <-> flat system-time scalars. The 7-octet CP56Time2a
// layout (IEC 60870-5-4): octets 0-1 = millisecond-of-day LE16,
// octet 2 = minute (bits 0..5) + SUC (bit6) + IV (bit7),
// octet 3 = hour (bits 0..4) + SU (bit7),
// octet 4 = day-of-week (bits 5..7) + day-of-month (bits 0..4),
// octet 5 = month (bits 0..3), octet 6 = year-1900 (bits 0..6) +
// IV2 (bit7). TwinCAT returns/accepts a TIMESTRUCT; here the
// fields are scalar outputs / inputs.
FUNCTION_BLOCK CP56Time2a_TO_SYSTEMTIME
VAR_INPUT
    pTime : ARRAY[0..6] OF BYTE;
END_VAR
VAR_OUTPUT
    nYear : UDINT;               // full year (1900 + field)
    nMonth : UDINT;              // 1..12
    nDay : UDINT;                // 1..31
    nHour : UDINT;               // 0..23
    nMinute : UDINT;             // 0..59
    nSecond : UDINT;             // 0..59
    nMs : UDINT;                 // 0..999
    bIV : BOOL;                  // invalid flag
    bSU : BOOL;                  // substituted / summer-time
END_VAR
VAR
    msod : UDINT;
END_VAR
    /* octets 0-1 = millisecond-of-minute LE16 (sec*1000+ms,
       max 59999); octet 2 = minute (bits 0..5) + SUC + IV */
    msod := (BYTE_TO_UDINT(pTime[0]) +
             BYTE_TO_UDINT(pTime[1]) * 256);
    nMs := msod MOD 1000;
    msod := msod / 1000;
    nSecond := msod MOD 60;
    nMinute := BYTE_TO_UDINT(pTime[2]) AND 16#3F;
    nHour := BYTE_TO_UDINT(pTime[3]) AND 16#1F;
    nDay := BYTE_TO_UDINT(pTime[4]) AND 16#1F;
    nMonth := BYTE_TO_UDINT(pTime[5]) AND 16#0F;
    nYear := 1900 + (BYTE_TO_UDINT(pTime[6]) AND 16#7F);
    bIV := (BYTE_TO_UDINT(pTime[2]) AND 16#80) <> 0;
    bSU := ((BYTE_TO_UDINT(pTime[2]) AND 16#40) <> 0) OR
           ((BYTE_TO_UDINT(pTime[3]) AND 16#80) <> 0);
END_FUNCTION_BLOCK

FUNCTION_BLOCK SYSTEMTIME_TO_CP56Time2a
VAR_INPUT
    nYear : UDINT;
    nMonth : UDINT;
    nDay : UDINT;
    nHour : UDINT;
    nMinute : UDINT;
    nSecond : UDINT;
    nMs : UDINT;
    bIV : BOOL;
    bSU : BOOL;
END_VAR
VAR_OUTPUT
    pTime : ARRAY[0..6] OF BYTE;
END_VAR
VAR
    msod : UDINT;
    y : UDINT;
END_VAR
    /* octets 0-1 = (sec*1000+ms) LE16, the ms-within-minute
       field (max 59999) */
    msod := nSecond * 1000 + nMs;
    pTime[0] := UDINT_TO_BYTE(msod MOD 256);
    pTime[1] := UDINT_TO_BYTE((msod / 256) MOD 256);
    pTime[2] := UDINT_TO_BYTE(nMinute AND 16#3F);
    IF bSU THEN pTime[2] := UDINT_TO_BYTE(BYTE_TO_UDINT(pTime[2]) OR 16#40); END_IF;
    IF bIV THEN pTime[2] := UDINT_TO_BYTE(BYTE_TO_UDINT(pTime[2]) OR 16#80); END_IF;
    pTime[3] := UDINT_TO_BYTE(nHour AND 16#1F);
    IF bSU THEN pTime[3] := UDINT_TO_BYTE(BYTE_TO_UDINT(pTime[3]) OR 16#80); END_IF;
    pTime[4] := UDINT_TO_BYTE(nDay AND 16#1F);
    pTime[5] := UDINT_TO_BYTE(nMonth AND 16#0F);
    y := nYear;
    IF y >= 1900 THEN y := y - 1900; END_IF;
    pTime[6] := UDINT_TO_BYTE(y AND 16#7F);
    IF bIV THEN pTime[6] := UDINT_TO_BYTE(BYTE_TO_UDINT(pTime[6]) OR 16#80); END_IF;
END_FUNCTION_BLOCK

// CP56Time2a_TO_CP24Time2a / CP56Time2a_TO_CP32Time2a — truncate
// the 7-octet CP56Time2a to the shorter CP24 (3 octets) /
// CP32 (4 octets) time tags.
FUNCTION_BLOCK CP56Time2a_TO_CP24Time2a
VAR_INPUT
    pIn : ARRAY[0..6] OF BYTE;
END_VAR
VAR_OUTPUT
    pOut : ARRAY[0..2] OF BYTE;
END_VAR
    pOut[0] := pIn[0];
    pOut[1] := pIn[1];
    pOut[2] := pIn[2];
END_FUNCTION_BLOCK

FUNCTION_BLOCK CP56Time2a_TO_CP32Time2a
VAR_INPUT
    pIn : ARRAY[0..6] OF BYTE;
END_VAR
VAR_OUTPUT
    pOut : ARRAY[0..3] OF BYTE;
END_VAR
    pOut[0] := pIn[0];
    pOut[1] := pIn[1];
    pOut[2] := pIn[2];
    pOut[3] := pIn[3];
END_FUNCTION_BLOCK

// F_iecGetSPI / F_iecSetSPI — single-point information bit
// (bit 0 of the 1-octet M_SP info element).
FUNCTION F_iecGetSPI : BOOL
VAR_INPUT
    nValue : UDINT;               // raw info element octet
END_VAR
    F_iecGetSPI := (nValue AND 16#01) <> 0;
END_FUNCTION

FUNCTION F_iecSetSPI : UDINT
VAR_INPUT
    nValue : UDINT;
    bSPI : BOOL;
END_VAR
    IF bSPI THEN
        F_iecSetSPI := (nValue AND 16#FE) OR 16#01;
    ELSE
        F_iecSetSPI := nValue AND 16#FE;
    END_IF
END_FUNCTION

// F_iecGetDPI / F_iecSetDPI — double-point information (bits 0..1:
// 0=off 1=on 2=indeterminate 3=off+on invalid).
FUNCTION F_iecGetDPI : UDINT
VAR_INPUT
    nValue : UDINT;
END_VAR
    F_iecGetDPI := nValue AND 16#03;
END_FUNCTION

FUNCTION F_iecSetDPI : UDINT
VAR_INPUT
    nValue : UDINT;
    nDPI : UDINT;
END_VAR
    F_iecSetDPI := (nValue AND 16#FC) OR (nDPI AND 16#03);
END_FUNCTION

// F_iecGetSCS / F_iecSetSCS — single-command state (C_SC select/
// execute state bits in the command response info element).
FUNCTION F_iecGetSCS : UDINT
VAR_INPUT
    nValue : UDINT;
END_VAR
    F_iecGetSCS := (nValue / 16) AND 16#03;
END_FUNCTION

FUNCTION F_iecSetSCS : UDINT
VAR_INPUT
    nValue : UDINT;
    nSCS : UDINT;
END_VAR
    F_iecSetSCS := (nValue AND 16#CF) OR ((nSCS AND 16#03) * 16);
END_FUNCTION

// F_iecGetDCS / F_iecSetDCS — double-command state (C_DC).
FUNCTION F_iecGetDCS : UDINT
VAR_INPUT
    nValue : UDINT;
END_VAR
    F_iecGetDCS := (nValue / 16) AND 16#03;
END_FUNCTION

FUNCTION F_iecSetDCS : UDINT
VAR_INPUT
    nValue : UDINT;
    nDCS : UDINT;
END_VAR
    F_iecSetDCS := (nValue AND 16#CF) OR ((nDCS AND 16#03) * 16);
END_FUNCTION

// F_iecGetQDS — quality-descriptor octet mask (bit7 IV, bit6 NT,
// bit5 SUC, bit4 BL, bit0 OV).
FUNCTION F_iecGetQDS : UDINT
VAR_INPUT
    nValue : UDINT;
END_VAR
    F_iecGetQDS := nValue AND 16#FF;
END_FUNCTION

FUNCTION F_iecSetQDS : UDINT
VAR_INPUT
    nValue : UDINT;
    nQDS : UDINT;
END_VAR
    F_iecSetQDS := (nValue AND 16#FF00) OR (nQDS AND 16#FF);
END_FUNCTION

// F_iecIncVTI / F_iecDecVTI — wrap-around increment/decrement of
// a 15-bit IEC sequence counter (sequence numbers mod 32768).
FUNCTION F_iecIncVTI : UDINT
VAR_INPUT
    nVTI : UDINT;
END_VAR
VAR
    v : UDINT;
END_VAR
    v := nVTI AND 16#7FFF;
    IF v >= 32767 THEN
        F_iecIncVTI := 0;
    ELSE
        F_iecIncVTI := v + 1;
    END_IF
END_FUNCTION

FUNCTION F_iecDecVTI : UDINT
VAR_INPUT
    nVTI : UDINT;
END_VAR
VAR
    v : UDINT;
END_VAR
    v := nVTI AND 16#7FFF;
    IF v = 0 THEN
        F_iecDecVTI := 32767;
    ELSE
        F_iecDecVTI := v - 1;
    END_IF
END_FUNCTION

// F_iecGetAOQuality / F_iecSetAOQuality / F_iecGetAOTimeTag /
// F_iecInitAOEntry — AO (application object) entry helpers on a
// flat UDINT slot: bits 8..15 quality, bits 0..15 time tag.
FUNCTION F_iecGetAOQuality : UDINT
VAR_INPUT
    nAO : UDINT;
END_VAR
    F_iecGetAOQuality := (nAO / 256) AND 16#FF;
END_FUNCTION

FUNCTION F_iecSetAOQuality : UDINT
VAR_INPUT
    nAO : UDINT;
    nQuality : UDINT;
END_VAR
    F_iecSetAOQuality := (nAO AND 16#FFFF00FF) OR
                         ((nQuality AND 16#FF) * 256);
END_FUNCTION

FUNCTION F_iecGetAOTimeTag : UDINT
VAR_INPUT
    nAO : UDINT;
END_VAR
    F_iecGetAOTimeTag := nAO AND 16#FFFF;
END_FUNCTION

FUNCTION F_iecInitAOEntry : UDINT
VAR_INPUT
    nAO : UDINT;
END_VAR
    F_iecInitAOEntry := nAO AND 16#FFFF0000;
END_FUNCTION

// Version function covering FB_GetIec870_Version-style queries.
FUNCTION GetIec870_Version : UDINT
    GetIec870_Version := 16#0100;   // v1.00
END_FUNCTION
